(* IEC 61131-3 sources: daoli-st-library/DL_Process (part 63) *)

(* ---- FB_DL_ChamberSeasoningTrack.st ---- *)
(*==============================================================================
 * 组件名称 (Component)  : FB_DL_ChamberSeasoningTrack
 * 所属子库 (Sublibrary) : DL_Process
 * 当前版本 (Version)    : 1.0.0
 * 组件分类 (Category)   : 功能块（FUNCTION_BLOCK）· 腔体 seasoning 台账与放行判定
 * 兼容性   (Platform)   : CODESYS 3.5 / TwinCAT 3 / 汇川 InoProShop / Schneider Machine Expert
 *                         仅依赖 Standard.library（R_TRIG / LEN / LEFT / ABS / MIN / MAX / LIMIT），零厂商方言
 * 接口依赖 (Depends)    : E_DL_Ne107Status —— 唯一属主为 DL_Device 子库的契约件
 *                         I_DL_DeviceHealth（R13 泳道 A1）。本文件只引用成员，不重定义枚举体。
 * 功能描述 (Function)   : seasoning（腔体调机）片数 + 膜厚台账 + 放行判定。每片完成后累计
 *                         片数、累计工艺时长、膜厚均值与趋势；**双判据**（片数达标 **且** 时长
 *                         达标）才放行；连续越窗自动降级 eNotReady；配方名只作标签与校验键。
 * 边界     (Boundary)   : ① **不做配方存储** —— sRecipeName 只作为标签与校验键传入，配方本体
 *                         归 FB_DL_RecipeManager；② **不做膜厚测量** —— 膜厚与均匀性由量测机台
 *                         引脚注入；③ 不做 SPC 判异（只做越窗计数与连续计数）；④ 不做 MES 上报。
 * 分层声明 (Layer)      : 工艺层（DL_Process）。零全局变量表引用、零外部变量声明、零物理 IO。
 * 段序     (Segments)   : 段1 实例无条件刷新 → 段2 复位通道（CASE 前，R39）→ 段3 配方标签闸门
 *                         （R37 显式截断）与参数钳位 → 段4 单片完成受理（R24/R25/R44）→
 *                         段5 状态机 → 段6 码位单一优先级链 → 段7 出口钳位与保持重写。
 * 枚举映射表 (R31)      : eIdle(0)→标签 0｜eTracking(10)→标签 10｜eQualified(20)→标签 20｜
 *                         eNotReady(30)→标签 30｜eFault(99)→标签 99。每个成员有且仅有一个
 *                         显式标签，ELSE 只接脏值（02FB）。
 * 单拍标志清单 (R25)    : bWaferDone —— 预清零点：段1 每拍被实例输出覆盖；置位点：段1
 *                         `_bWaferReq := _fbTrigWafer.Q AND (NOT _bWaferConsumed)`；自清点：
 *                         段4 消费时置 `_bWaferConsumed := TRUE`，bWaferDone 回 FALSE 即解除。
 *                         bReset —— 预清零点：段1 覆盖 _bResetEdge；置位点：段1 实例调用；
 *                         自清点：紧随实例调用的 _bResetEdge 赋值行。
 * 保持位清单 (R27)      : bRelease 逐拍由 _bReleaseLatched 重写；eQualify 逐拍由 _eState 映射；
 *                         nCount / nNgCount / tAccum / fThickAvg / fThickSlope 逐拍由内部
 *                         台账量重写并夹域。复位沿清台账并递增轮次号。
 * 定时器清单 (R40)      : 无 TON/TOF 实例。工艺时长由引脚 tProcessTime 累加（台账语义），
 *                         不存在跨段恒真的定时输入；片数与时长的「达标」判据均为纯比较式。
 * 三元一致表 (R35)      : 片数目标守卫 1~10000 / 封顶 10000 / 判据 `>=`｜
 *                         连续越窗阈守卫 1~10 / 封顶 10 / 判据 `>=`｜
 *                         膜厚容差守卫 0.5~50 % / 封顶 50 / 判据 `>`（越窗）。
 * 镜像量清单 (R38)      : sRecipeName 的长度经 LEN 一次锁存为 _nNameLen，截断判定与登记
 *                         全部读该锁存量，绝不二次取长度；fThickness 与 fUniformity 在段4
 *                         单次锁存后参与全部判据。
 * 开源溯源 (Origin)     : 原创实现（参考 SEMI/半导体厂务公开的 seasoning 台账惯例，以及
 *                         ISA-88 公开的批次/相语义，T2-8 只借「批次台账 + 放行」的组织形态；
 *                         配方名仅作标签、台账只做累计与双判据）。ISA-88 为公开标准条款，
 *                         不声称「符合 ISA-88」；实现、码位、引脚契约 100% 本库独立设计，
 *                         clean-room 编写，未复制任何源码行。许可证说明：无代码借鉴对象，
 *                         本文件为本库原创，随本库许可证发布。
 * 验收向量 (Acceptance) :
 *   V1 25 片、每片 24 min、膜厚 100 ± 2 nm（目标 100、容差 5 %）→ tAccum = 10 h、
 *      eQualified、bRelease = TRUE。
 *   V2（双判据）25 片但每片 10 min（总 4.17 h < 10 h）→ 16#0005_01CD、仍 eTracking、
 *      bRelease = FALSE。
 *   V3（V-A 缺失键）sRecipeName = '' → 16#0005_02F9 锁存、bRelease 强制 FALSE
 *      （安全侧：台账不可信不得放行）。
 *   V4（V-B 串上限，R37）sRecipeName 传 40 字符（超 STRING(32)）→ 入口判 LEN 后置
 *      16#0005_01CE，按截断后的名字登记台账，**不得**依赖赋值隐式截断后静默使用。
 *   V5（V-D 复位首拍）bReset 后 nCount = 0、tAccum = T#0S、nRoundId + 1、bRelease = FALSE；
 *      **不得**保留上一轮 fThickSlope 的首片基准（R41：恢复不重头）。
 * 偏离留档 (Deviation)  :
 *   ① sRecipeName 引脚类型由 STRING(32) 提升为 STRING(80)：若按 STRING(32) 声明，超长截断
 *      会发生在**调用方赋值**那一行，本件永远看不到长度越限，01CE 成为死码 —— 这正是 R37
 *      要消灭的「静默截断」。提升到 STRING(80) 后由本件判 LEN、显式置码、按截断名登记，
 *      登记缓冲仍为 STRING(32)（_sRecipeTag），行为与规格 V4 一致。
 *   ② 工艺时长用 tProcessTime 累加而非墙钟：一台上位机可能同时跟踪多条腔体，墙钟会把
 *      「等待/待机」算进 seasoning 时长；引脚注入的工艺耗时才是台账口径。
 *   ③ 越窗判据取「膜厚相对偏差 > fThickTol 或 均匀性 > fUnifLimit」的**并集**：均匀性越限
 *      同样是「膜质未稳」的证据，只盯膜厚会漏掉「厚度对但均匀性崩」的片子。
 *   ④ 量测值非有限/越域并入 16#0005_02FA：规格故障表只给三个码，量测值不可信属于
 *      「台账数据源坏了」，与计数溢出同属「台账不可继续累加」的语义，故共用该码；
 *      不发生任何累加（本片不入账），也不会放行。
 * 修订历史 (Revision)   :
 *   2026-11-15  v1.0.0  首版入库（Round 13 · 泳道 C · DL_Process 第 25 件）
 *============================================================================*)

(*-----------------------------------------------------------------------------
 * 枚举: E_DL_SeasonState（归属 FB_DL_ChamberSeasoningTrack，同文件发布）
 *----------------------------------------------------------------------------*)
TYPE E_DL_SeasonState :
(
    eIdle      := 0,    // 空闲：未使能或参数未就绪 / Idle, disabled or parameters not ready
    eTracking  := 10,   // 台账中：逐片累计，双判据未齐 / Tracking, accumulating wafers
    eQualified := 20,   // 已放行：片数与时长双达标 / Qualified, both criteria met
    eNotReady  := 30,   // 不具备放行条件：连续越窗降级 / Not ready, consecutive out-of-window wafers
    eFault     := 99    // 故障：配方键缺失或计数溢出 / Fault, missing recipe key or counter overflow
) UINT;
END_TYPE

FUNCTION_BLOCK FB_DL_ChamberSeasoningTrack
VAR_INPUT
    bEnable       : BOOL;                   // 使能（Enable），FALSE = 冻结台账与放行；复位通道不受其屏蔽 / Enable, FALSE freezes the ledger
    bReset        : BOOL;                   // 复位（Reset），上升沿清台账并重开新一轮 / Rising edge clears the ledger and opens a new round
    bWaferDone    : BOOL;                   // 单片完成（One-shot wafer done），上升沿受理（R24）/ One-shot wafer done, rising edge only
    fThickness    : REAL;                   // 本片膜厚（Wafer thickness）[nm]，域 0~10000 / Wafer thickness [nm], 0 to 10000
    fUniformity   : REAL;                   // 本片均匀性（Uniformity）[%]，域 0~100 / Uniformity [%], 0 to 100
    sRecipeName   : STRING(80);             // 配方名标签（Recipe tag），域非空，超 32 字符显式截断并置码（偏离留档①）/ Recipe tag, truncated explicitly
    fThickTarget  : REAL;                   // 膜厚目标（Thickness target）[nm]，域 >0 / Thickness target [nm], must be positive
    fThickTol     : REAL := 5.0;            // 膜厚相对容差（Thickness tolerance）[%]，域 0.5~50，默认 5.0 / Thickness tolerance [%]
    fUnifLimit    : REAL := 3.0;            // 均匀性上限（Uniformity limit）[%]，域 0.1~20，默认 3.0 / Uniformity limit [%]
    nCountTarget  : INT := 25;              // 片数目标（Wafer count target）[片]，域 1~10000，默认 25 / Wafer count target [pcs]
    tTimeTarget   : TIME := T#10H;          // 工艺时长目标（Process time target），域 1 min~1000 h，默认 10 h / Process time target
    nConsecNgLimit : INT := 2;              // 连续越窗降级阈值（Consecutive out-of-window limit）[片]，域 1~10，默认 2 / Consecutive limit [pcs]
    tProcessTime  : TIME;                   // 本片工艺耗时（Process time of this wafer），由上层引脚注入 / Process time injected by the caller
END_VAR

VAR_OUTPUT
    nCount        : INT;                    // 已 seasoning 片数（Seasoned wafer count）[片]，逐拍重写 / Seasoned wafer count [pcs]
    nNgCount      : INT;                    // 越窗片数（Out-of-window wafer count）[片]，逐拍重写 / Out-of-window wafer count [pcs]
    tAccum        : TIME;                   // 累计工艺时长（Accumulated process time），逐拍重写 / Accumulated process time
    fThickAvg     : REAL;                   // 膜厚均值（Mean thickness）[nm]，逐拍重写 / Mean thickness [nm]
    fThickSlope   : REAL;                   // 膜厚趋势（Thickness trend）[nm/片]，首末差除以片数差 / Thickness trend [nm/pc]
    bRelease      : BOOL;                   // 放行（Release），保持语义（R27）/ Release, held
    eQualify      : E_DL_SeasonState;       // 判定状态（Qualification state），逐拍重写 / Qualification state
    nRoundId      : UINT;                   // 本轮编号（Round id），复位递增，供 MES 对齐 / Round id, incremented on reset
    eHealth       : E_DL_Ne107Status;       // 健康态（NE107 health），引用属主 A1 的枚举 / NE107 health, owned by A1
    uDiagCode     : UDINT;                  // 诊断码（Diagnostic code），本拍单一优先级链输出 / Diagnostic code, single priority chain
    uErrorId      : UDINT;                  // 故障码（Error code），仅故障级码，0 = 无故障 / Fault-level code, 0 = no fault
    bError        : BOOL;                   // 故障标志（Error），仅故障级码置位 / TRUE only for fault-level codes
END_VAR

VAR
    _eState       : E_DL_SeasonState := E_DL_SeasonState.eIdle;    // 内部状态（Internal state）/ Internal state value
    _bWaferReq    : BOOL;                   // 单片完成单拍请求（Wafer done request）/ Wafer done one-shot request
    _bWaferConsumed : BOOL;                 // 单片完成已消费（Wafer consumed flag）/ Wafer consumed flag
    _bResetEdge   : BOOL;                   // 复位沿单拍标志（Reset one-shot flag）/ Reset one-shot flag
    _uFaultCode   : UDINT;                  // 本拍故障级码（Fault-level code this scan）/ Fault-level code of this scan
    _uFaultLatched : UDINT;                 // 故障码锁存（Latched fault code），仅复位清除 / Latched fault code, reset only
    _uInfoCode    : UDINT;                  // 本拍信息级码（Info-level code this scan）/ Info-level code of this scan
    _bFaultCond   : BOOL;                   // 故障条件（Fault condition）/ Fault condition flag
    _sRecipeTag   : STRING(32);             // 台账登记的配方标签（Registered recipe tag），截断后 32 字符 / Recipe tag after truncation
    _nNameLen     : INT;                    // 配方名长度（Recipe name length）[字符]，一次锁存（R38）/ Recipe name length, latched once
    _bTruncFlag   : BOOL;                   // 截断发生标志（Truncation flag），R37 显式置位 / Truncation flag, set explicitly (R37)
    _bKeyOk       : BOOL;                   // 配方键与目标合法（Key and target valid）/ Key and target valid
    _fThickSnap   : REAL;                   // 膜厚快照（Thickness snapshot）[nm]，单次锁存 / Thickness snapshot [nm]
    _fUnifSnap    : REAL;                   // 均匀性快照（Uniformity snapshot）[%]，单次锁存 / Uniformity snapshot [%]
    _fTolEff      : REAL;                   // 生效膜厚容差（Effective thickness tolerance）[%] / Effective thickness tolerance [%]
    _fUnifLimEff  : REAL;                   // 生效均匀性上限（Effective uniformity limit）[%] / Effective uniformity limit [%]
    _nCountTgtEff : INT;                    // 生效片数目标（Effective count target）[片] / Effective count target [pcs]
    _nConsecEff   : INT;                    // 生效连续越窗阈（Effective consecutive limit）[片] / Effective consecutive limit [pcs]
    _tTimeTgtEff  : TIME;                   // 生效时长目标（Effective time target）/ Effective time target
    _nCountInt    : INT;                    // 内部片数台账（Internal wafer count）[片] / Internal wafer count [pcs]
    _nNgInt       : INT;                    // 内部越窗片数（Internal out-of-window count）[片] / Internal out-of-window count [pcs]
    _nConsecNg    : INT;                    // 当前连续越窗片数（Current consecutive out-of-window count）[片] / Current consecutive count [pcs]
    _tAccumInt    : TIME;                   // 内部累计时长（Internal accumulated time）/ Internal accumulated time
    _fThickSum    : REAL;                   // 膜厚累加（Thickness sum）[nm] / Thickness sum [nm]
    _fThickFirst  : REAL;                   // 首片膜厚（First wafer thickness）[nm]，趋势基准 / First wafer thickness [nm]
    _fThickLast   : REAL;                   // 末片膜厚（Last wafer thickness）[nm] / Last wafer thickness [nm]
    _bFirstSet    : BOOL;                   // 首片基准已装（First sample recorded）/ First sample recorded flag
    _fDevPct      : REAL;                   // 膜厚相对偏差（Relative thickness deviation）[%] / Relative thickness deviation [%]
    _bOutWin      : BOOL;                   // 本片越窗（Out of window this wafer）/ Out of window this wafer
    _bReleaseLatched : BOOL;                // 放行锁存（Release latch），复位清除 / Release latch, reset only
    _nRoundIdInt  : UINT;                   // 内部轮次号（Internal round id），复位递增 / Internal round id, incremented on reset
    _bCountOk     : BOOL;                   // 片数达标（Count criterion met）/ Count criterion met
    _bTimeOk      : BOOL;                   // 时长达标（Time criterion met）/ Time criterion met
    _fbTrigWafer  : R_TRIG;                 // 单片完成上升沿（Wafer done rising edge）/ Wafer done rising edge
    _fbTrigReset  : R_TRIG;                 // 复位上升沿（Reset rising edge）/ Reset rising edge
END_VAR

VAR CONSTANT
    DL_SEA_NAME_MAX   : INT  := 32;          // 配方标签登记宽度（Registered tag width）[字符]，与 STRING(32) 一致 / Registered tag width
    DL_SEA_REAL_MAX   : REAL := 3.4E38;      // 单精度有限值判据幅值（Finite magnitude bound）/ Finite bound for REAL inputs
    DL_SEA_EPS        : REAL := 1.0E-6;      // 浮点防零容差（Divide-guard epsilon）/ Float divide-guard epsilon
    DL_SEA_THICK_MAX  : REAL := 10000.0;     // 膜厚输入域上限（Thickness input bound）[nm] / Thickness input bound [nm]
    DL_SEA_UNIF_MAX   : REAL := 100.0;       // 均匀性输入域上限（Uniformity input bound）[%] / Uniformity input bound [%]
    DL_SEA_TOL_LO     : REAL := 0.5;         // 膜厚容差下限（Tolerance lower clamp）[%] / Tolerance lower clamp [%]
    DL_SEA_TOL_HI     : REAL := 50.0;        // 膜厚容差上限（Tolerance upper clamp）[%] / Tolerance upper clamp [%]
    DL_SEA_UNIFL_LO   : REAL := 0.1;         // 均匀性上限下限（Uniformity limit lower clamp）[%] / Uniformity lower clamp [%]
    DL_SEA_UNIFL_HI   : REAL := 20.0;        // 均匀性上限上限（Uniformity limit upper clamp）[%] / Uniformity upper clamp [%]
    DL_SEA_CNT_LO     : INT  := 1;           // 片数目标下限（Count target lower clamp）[片] / Count target lower clamp [pcs]
    DL_SEA_CNT_HI     : INT  := 10000;       // 片数目标上限（Count target upper clamp）[片] / Count target upper clamp [pcs]
    DL_SEA_CONS_LO    : INT  := 1;           // 连续阈下限（Consecutive limit lower clamp）[片] / Consecutive limit lower clamp [pcs]
    DL_SEA_CONS_HI    : INT  := 10;                 // 连续阈上限（Consecutive limit upper clamp）[片] / Consecutive limit upper clamp [pcs]
    DL_SEA_CNT_OVF    : INT  := 30000;       // 片数台账溢出阈（Count overflow threshold）[片] / Count overflow threshold [pcs]
    DL_SEA_TIME_OVF   : TIME := T#40D;       // 时长台账溢出阈（Time overflow threshold）[ms] / Time overflow threshold
    DL_SEA_TIME_MIN   : TIME := T#1M;        // 时长目标下限（Time target lower clamp）/ Time target lower clamp
    DL_SEA_TIME_MAX   : TIME := T#1000H;     // 时长目标上限（Time target upper clamp）/ Time target upper clamp
    DL_SEA_PCT        : REAL := 100.0;       // 百分比换算（Percent scale）[-] / Percent scale
    DL_SEA_ERR_KEY    : UDINT := 16#0005_02F9; // 0005_02F9 配方名为空或膜厚目标非正【故障级】/ Missing recipe or target, fault level
    DL_SEA_ERR_OVF    : UDINT := 16#0005_02FA; // 0005_02FA 片数或时长台账溢出【故障级】/ Counter overflow, fault level
    DL_SEA_ERR_STATE  : UDINT := 16#0005_02FB; // 0005_02FB 非法状态兜底【故障级】/ Illegal state fallback, fault level
    DL_SEA_INFO_SINGLE : UDINT := 16#0005_01CB; // 0005_01CB 单片越窗但未连续【信息级】/ Single out-of-window wafer, info level
    DL_SEA_INFO_CONS  : UDINT := 16#0005_01CC; // 0005_01CC 连续越窗达阈值降级【信息级】/ Consecutive limit reached, info level
    DL_SEA_INFO_TIME  : UDINT := 16#0005_01CD; // 0005_01CD 片数达标但时长未达标【信息级】/ Count reached, time pending, info level
    DL_SEA_INFO_TRUNC : UDINT := 16#0005_01CE; // 0005_01CE 配方名超 32 字符已显式截断【信息级】/ Recipe tag truncated explicitly, info level
END_VAR

// ============================================================================
// 段 1｜实例无条件周期刷新（R7/0.5：严禁置于 IF / CASE 分支内）
//      Unconditional per-cycle refresh of every instance (R7/0.5)
// ============================================================================
_fbTrigWafer(CLK := bWaferDone);                // 单片完成上升沿（Wafer done rising edge）
_bWaferReq := _fbTrigWafer.Q AND (NOT _bWaferConsumed);    // 单拍请求（R25 置位点）
_fbTrigReset(CLK := bReset);                    // 复位上升沿（Reset rising edge）
_bResetEdge := _fbTrigReset.Q;                  // 复位单拍标志紧随实例赋值（R25 自清点）

// 本拍码与条件预置（每拍重算；故障码以上拍锁存续用）
// Per-scan preset of codes and conditions, the fault code is carried from the latch
_uFaultCode := _uFaultLatched;                  // 故障码续用（Carry the latched fault code）
_uInfoCode  := 16#0000_0000;                    // 信息级码预清零（Info code preset to zero）
_bFaultCond := FALSE;                           // 故障条件预清零（Fault condition preset FALSE）
_bKeyOk     := FALSE;                           // 配方键闸门预置未通过（Key gate preset closed）
_bOutWin    := FALSE;                           // 越窗标志预置假（Out-of-window preset FALSE）

// 单片完成消费标志解除：输入回落即允许下一片（R25 生命周期闭环）
// Release the wafer consumption flag once the input falls
IF NOT bWaferDone THEN
    _bWaferConsumed := FALSE;                   // 允许下一次上升沿（Next rising edge accepted）
END_IF

// ============================================================================
// 段 2｜复位通道（R39：置于 CASE 之前，且不被掉使能分支屏蔽）
//      Reset path, before CASE and never masked by the disable branch
// ============================================================================
IF _bResetEdge THEN
    _nCountInt    := 0;                         // 片数台账清零（Wafer count cleared）
    _nNgInt       := 0;                         // 越窗片数清零（Out-of-window count cleared）
    _nConsecNg    := 0;                         // 连续越窗计数清零（Consecutive count cleared）
    _tAccumInt    := T#0S;                      // 累计时长清零（Accumulated time cleared）
    _fThickSum    := 0.0;                       // 膜厚累加清零（Thickness sum cleared）
    _fThickFirst  := 0.0;                       // 首片基准清除（First-sample basis cleared）
    _fThickLast   := 0.0;                       // 末片值清除（Last-sample value cleared）
    _bFirstSet    := FALSE;                     // 首片基准标志清除（First-sample flag cleared，R41）
    _bReleaseLatched := FALSE;                  // 放行锁存清除（Release latch cleared）
    _bTruncFlag   := FALSE;                     // 截断标志清除（Truncation flag cleared）
    _nRoundIdInt  := _nRoundIdInt + UINT#1;     // 轮次递增进位（Round id incremented）
    _uFaultLatched := 16#0000_0000;             // 故障码锁存清除（Latched fault code cleared）
    _uFaultCode   := 16#0000_0000;              // 本拍故障码清空，防止段6 重新锁存旧码（Clear this scan code）
    IF _eState = E_DL_SeasonState.eFault THEN
        _eState := E_DL_SeasonState.eIdle;      // 故障态回空闲（Fault state back to idle）
        _bFaultCond := FALSE;                   // 故障条件清除（Fault condition cleared）
    ELSIF _eState = E_DL_SeasonState.eQualified THEN
        _eState := E_DL_SeasonState.eTracking;  // 已放行轮次复位后重开台账（New round after a qualified round）
    ELSIF _eState = E_DL_SeasonState.eNotReady THEN
        _eState := E_DL_SeasonState.eTracking;  // 降级轮次复位后重开台账（New round after a degraded round）
    END_IF
END_IF

// ============================================================================
// 段 3｜配方标签闸门（R37：先判长度、显式置码、按截断名登记）与参数钳位
//      Recipe tag gate: length first, explicit code, then register the truncated tag
// ============================================================================
_nNameLen := LEN(sRecipeName);                  // 长度一次锁存（R38：此后全部判据读该值）
IF _nNameLen > DL_SEA_NAME_MAX THEN
    _sRecipeTag := LEFT(sRecipeName, DL_SEA_NAME_MAX);   // 按宽度取前缀后写回登记缓冲（预判后写，非回夹）
    _bTruncFlag := TRUE;                        // 截断标志显式置位（R37 核心：不静默）
    _uInfoCode  := DL_SEA_INFO_TRUNC;           // 0005_01CE 配方名超长已截断【信息级】/ Recipe tag truncated
ELSE
    _sRecipeTag := sRecipeName;                 // 未超长按原名登记（Register the tag as-is）
END_IF

IF _nNameLen = 0 THEN
    _bFaultCond := TRUE;                        // 配方键缺失（Missing recipe key）
    _uFaultCode := DL_SEA_ERR_KEY;              // 0005_02F9 配方名为空【故障级】/ Missing recipe, fault level
ELSIF (NOT (fThickTarget >= DL_SEA_EPS)) OR (fThickTarget > DL_SEA_THICK_MAX) THEN
    _bFaultCond := TRUE;                        // 膜厚目标非正或越域（Target not positive or out of domain）
    _uFaultCode := DL_SEA_ERR_KEY;              // 0005_02F9 膜厚目标非法【故障级】/ Illegal target, fault level
ELSE
    _bKeyOk := TRUE;                            // 键与目标合法（Key and target valid）
END_IF

// 参数域钳位（R35：守卫、封顶与判据同向）
// Parameter clamping so that guard, ceiling and comparison stay in step (R35)
_fTolEff      := LIMIT(DL_SEA_TOL_LO, fThickTol, DL_SEA_TOL_HI);            // 膜厚容差 0.5~50 %（Tolerance clamped）
_fUnifLimEff  := LIMIT(DL_SEA_UNIFL_LO, fUnifLimit, DL_SEA_UNIFL_HI);       // 均匀性上限 0.1~20 %（Uniformity limit clamped）
_nCountTgtEff := LIMIT(DL_SEA_CNT_LO, nCountTarget, DL_SEA_CNT_HI);         // 片数目标 1~10000（Count target clamped）
_nConsecEff   := LIMIT(DL_SEA_CONS_LO, nConsecNgLimit, DL_SEA_CONS_HI);     // 连续阈 1~10（Consecutive limit clamped）
_tTimeTgtEff := tTimeTarget;                    // 时长目标取引脚值（Time target taken from the pin）
IF _tTimeTgtEff < DL_SEA_TIME_MIN THEN
    _tTimeTgtEff := DL_SEA_TIME_MIN;            // 时长目标下限钳位（Time target lower clamp）
ELSIF _tTimeTgtEff > DL_SEA_TIME_MAX THEN
    _tTimeTgtEff := DL_SEA_TIME_MAX;            // 时长目标上限钳位（Time target upper clamp）
END_IF

// ============================================================================
// 段 4｜单片完成受理（R24/R25；R44 清码点绑定新片起点）
//      Wafer completion acceptance, info codes cleared at each wafer start (R44)
// ============================================================================
IF _bWaferReq AND (NOT _bWaferConsumed) AND (_eState = E_DL_SeasonState.eTracking) AND _bKeyOk THEN
    _bWaferConsumed := TRUE;                    // 消费单片沿（Wafer edge consumed）
    _uInfoCode      := 16#0000_0000;            // 新片起点清信息码（R44：清码点绑定新片起点）
    _fThickSnap     := fThickness;              // 膜厚快照（Thickness snapshot）
    _fUnifSnap      := fUniformity;             // 均匀性快照（Uniformity snapshot）

    IF (NOT (_fThickSnap >= 0.0 AND _fThickSnap <= DL_SEA_THICK_MAX))
    OR (NOT (_fUnifSnap >= 0.0 AND _fUnifSnap <= DL_SEA_UNIF_MAX)) THEN
        _bFaultCond := TRUE;                    // 量测值非有限或越域（Non-finite or out-of-domain measurement）
        _uFaultCode := DL_SEA_ERR_OVF;          // 0005_02FA 量测值非法并入溢出码【故障级】/ Illegal measurement folded in
    ELSE
        _nCountInt := _nCountInt + 1;           // 片数 +1（Wafer counted）
        _fThickSum := _fThickSum + _fThickSnap; // 膜厚累加（Thickness accumulated）
        _fThickLast := _fThickSnap;             // 末片膜厚（Last wafer thickness）
        IF NOT _bFirstSet THEN
            _fThickFirst := _fThickSnap;        // 首片基准只在首片装一次（First-sample basis once）
            _bFirstSet   := TRUE;               // 基准已装（Basis recorded）
        END_IF
        _tAccumInt := _tAccumInt + tProcessTime;    // 累计工艺时长（Process time accumulated）

        // 越窗判据：膜厚相对偏差 或 均匀性越限（偏离留档③）
        //     Out-of-window when the thickness deviation or the uniformity exceeds its limit
        _fDevPct := ABS(_fThickSnap - fThickTarget) / fThickTarget * DL_SEA_PCT;    // 相对偏差（Relative deviation）
        IF (_fDevPct > _fTolEff) OR (_fUnifSnap > _fUnifLimEff) THEN
            _bOutWin := TRUE;                   // 本片越窗（Out of window）
        END_IF

        IF _bOutWin THEN
            _nNgInt    := _nNgInt + 1;          // 越窗片数 +1（Out-of-window counted）
            _nConsecNg := _nConsecNg + 1;       // 连续越窗 +1（Consecutive count increments）
            IF _nConsecNg >= _nConsecEff THEN
                _uInfoCode := DL_SEA_INFO_CONS; // 0005_01CC 连续越窗达阈值降级【信息级】/ Consecutive limit reached
            ELSE
                _uInfoCode := DL_SEA_INFO_SINGLE;   // 0005_01CB 单片越窗但未连续【信息级】/ Single out-of-window wafer
            END_IF
        ELSE
            _nConsecNg := 0;                    // 未越窗则连续计数清零（Consecutive count resets）
        END_IF

        // 台账溢出守卫（R35：守卫 30000 片 / 40 天，判据 >=）
        //     Ledger overflow guard
        IF (_nCountInt >= DL_SEA_CNT_OVF) OR (_tAccumInt >= DL_SEA_TIME_OVF) THEN
            _bFaultCond := TRUE;                // 台账溢出（Ledger overflow）
            _uFaultCode := DL_SEA_ERR_OVF;      // 0005_02FA 台账溢出【故障级】/ Ledger overflow, fault level
        END_IF
    END_IF
END_IF

// 双判据（片数达标 且 时长达标）：片数达标而时长未达标时只给信息码，不放行
// Dual criteria: the count alone never releases the chamber
_bCountOk := _nCountInt >= _nCountTgtEff;       // 片数判据（Count criterion）
_bTimeOk  := _tAccumInt >= _tTimeTgtEff;        // 时长判据（Time criterion）
IF _bCountOk AND (NOT _bTimeOk) THEN
    _uInfoCode := DL_SEA_INFO_TIME;             // 0005_01CD 片数达标但时长未达标【信息级】/ Count reached, time pending
END_IF

// ============================================================================
// 段 5｜状态机（ENUM + CASE，含 ELSE 非法状态兜底）
//      State machine with an explicit ELSE fallback
// ============================================================================
IF _bFaultCond THEN
    _bReleaseLatched := FALSE;                  // 安全侧：台账不可信时强制撤销放行（Safety: release revoked on any fault）
    _eState := E_DL_SeasonState.eFault;         // 故障条件优先于状态机（Fault outranks the machine）
END_IF

// 掉使能冻结分支：显式排除故障态（R39 合法写法①），复位通道仍可从故障态退出
// Disable branch explicitly excludes the fault state so the reset path still works
IF (NOT bEnable) AND (_eState <> E_DL_SeasonState.eFault) THEN
    _eState := E_DL_SeasonState.eIdle;          // 冻结回空闲（Freeze back to idle）
END_IF

CASE _eState OF

    E_DL_SeasonState.eIdle: // 空闲：等键与目标就绪
        IF bEnable AND _bKeyOk AND (NOT _bFaultCond) THEN
            _eState := E_DL_SeasonState.eTracking;  // 门票就绪进台账（Enter tracking）
        END_IF

    E_DL_SeasonState.eTracking: // 台账中：双判据 / 连续越窗降级
        IF _bCountOk AND _bTimeOk THEN
            _bReleaseLatched := TRUE;           // 双判据齐：放行（Releases the chamber）
            _eState := E_DL_SeasonState.eQualified; // 进已放行（Enter qualified）
        ELSIF _nConsecNg >= _nConsecEff THEN
            _bReleaseLatched := FALSE;          // 降级：撤销放行（Degraded, release revoked）
            _eState := E_DL_SeasonState.eNotReady;  // 进不具备放行条件（Enter not ready）
        END_IF

    E_DL_SeasonState.eQualified: // 已放行：结论逐拍在段7 重写（R27），本分支只保留标签
        // 结论保持由段7 逐拍重写承担，此处保留空标签与原因注释（R31）
        // The held verdict is rewritten in segment 7, so this label stays empty (R31)

    E_DL_SeasonState.eNotReady: // 不具备放行条件：等复位重开一轮
        // 复位通道位于 CASE 之前（段2），此处保留空标签与原因注释（R31/R41）
        // Reset happens in segment 2, so this label stays empty (R31/R41)

    E_DL_SeasonState.eFault: // 故障：等复位沿（段2）
        // 复位通道位于 CASE 之前，此分支无需动作（R39）
        // The reset path sits before CASE, so no action is needed here (R39)

    ELSE // 兜底：非法状态
        _uFaultCode := DL_SEA_ERR_STATE;        // 0005_02FB 非法状态兜底【故障级】/ Illegal state fallback
        _bFaultCond := TRUE;                    // 置故障条件（Raise the fault condition）
        _eState     := E_DL_SeasonState.eFault; // 强制回故障态（Force the fault state）
END_CASE

// ============================================================================
// 段 6｜码位单一优先级链（全拍只写一次，信息级不置 bError）
//      Single priority chain for the codes, written once per scan
// ============================================================================
IF _uFaultCode <> 16#0000_0000 THEN
    _uFaultLatched := _uFaultCode;              // 故障码锁存（Latched until reset）
    uErrorId  := _uFaultCode;                   // 故障级码优先（Fault-level code wins）
    uDiagCode := _uFaultCode;                   // 诊断码同源（Diagnostic code mirrors the fault）
    bError    := TRUE;                          // 故障标志置位（Error flag raised）
ELSIF _uInfoCode <> 16#0000_0000 THEN
    uErrorId  := 16#0000_0000;                  // 信息级不占故障码（Info level leaves the fault code empty）
    uDiagCode := _uInfoCode;                    // 诊断码取信息级码（Diagnostic code takes the info code）
    bError    := FALSE;                         // 信息级不置故障位（Info level never raises the error flag）
ELSE
    uErrorId  := 16#0000_0000;                  // 无码（No code）
    uDiagCode := 16#0000_0000;                  // 无码（No code）
    bError    := FALSE;                         // 无故障（No error）
END_IF

// ============================================================================
// 段 7｜出口钳位与保持语义重写（R27/R43；台账量逐拍重写，绝不靠进入那一拍）
//      Output clamping and held-semantics rewrite (R27/R43)
// ============================================================================
nCount    := LIMIT(0, _nCountInt, DL_SEA_CNT_OVF);      // 片数夹进 0~30000（Count clamped）
nNgCount  := LIMIT(0, _nNgInt, DL_SEA_CNT_OVF);         // 越窗片数夹进 0~30000（Out-of-window clamped）
tAccum    := _tAccumInt;                                // 累计时长逐拍重写（Accumulated time rewritten）
IF _nCountInt > 0 THEN
    fThickAvg := _fThickSum / INT_TO_REAL(_nCountInt);  // 膜厚均值（Mean thickness），除零已由计数守卫
ELSE
    fThickAvg := 0.0;                                   // 无片时均值 0（Zero mean without wafers）
END_IF
IF (_nCountInt >= 2) AND _bFirstSet THEN
    fThickSlope := (_fThickLast - _fThickFirst) / INT_TO_REAL(_nCountInt - 1);  // 首末差/片数差（Trend per wafer）
ELSE
    fThickSlope := 0.0;                                 // 单片或未装基准时趋势 0（Zero trend before a basis exists）
END_IF
bRelease  := _bReleaseLatched;                          // 放行逐拍重写（Release rewritten every scan）
eQualify  := _eState;                                   // 判定状态逐拍重写（Qualification state rewritten）
nRoundId  := _nRoundIdInt;                              // 轮次号逐拍重写（Round id rewritten every scan）

// 健康态仲裁（引用属主 A1 的四态语言）
// Health arbitration mapped onto the A1 health language
IF _eState = E_DL_SeasonState.eFault THEN
    eHealth := E_DL_Ne107Status.eFailure;       // 故障：台账不可信（Failure）
ELSIF NOT bEnable THEN
    eHealth := E_DL_Ne107Status.eUnknown;       // 未知：未使能（Unknown）
ELSIF _eState = E_DL_SeasonState.eNotReady THEN
    eHealth := E_DL_Ne107Status.eMaintenanceReq;    // 需维护：连续越窗，需重新调机（Maintenance required）
ELSIF _bTruncFlag THEN
    eHealth := E_DL_Ne107Status.eOutOfSpec;     // 越规：配方键被截断，台账对齐风险（Out of spec）
ELSIF _eState = E_DL_SeasonState.eQualified THEN
    eHealth := E_DL_Ne107Status.eOk;            // 正常：已放行（OK, released）
ELSE
    eHealth := E_DL_Ne107Status.eOk;            // 正常：台账进行中（OK, tracking）
END_IF

END_FUNCTION_BLOCK

(* ---- FB_DL_CipCleaningSeq.st ---- *)
(*==============================================================================
 * 组件名称 (Component)  : FB_DL_CipCleaningSeq
 * 所属子库 (Sublibrary) : DL_Process
 * 当前版本 (Version)    : 1.0.1
 * 兼容性 (Platform)   : CODESYS 3.5 / TwinCAT 3 / 汇川 InoProShop / Machine Expert
 *                         仅依赖 Standard.library（TON / R_TRIG），零厂商方言
 * 分类     (Category)   : 工艺段功能块（Function Block · CIP 原位清洗六相顺控）
 * 功能简述 (Function)   : CIP 原位清洗六相顺控：预冲洗 → 碱洗 → 中间冲洗 →
 *                         酸洗 → 终冲洗 → 消毒。核心纪律：相位计时受 TACT 联
 *                         锁暂停（温度/电导率/流量不达标不计时）；终冲洗以回
 *                         液电导率判终点（最长延时兜底）；回路就绪门控；换相
 *                         停泵间隔防混液；中止即排空隔离并失去清洁许可；偏差
 *                         计数供审计。本块不实现阀门矩阵/混流防护的物理设计
 *                         （属机械与管路设计），仅做就绪门控与指令编排。
 * 首扫说明 (Init note)  : 顺序型组件但全部状态由指令沿/电平驱动，免首扫
 *                         （R23/公约 0.1），无 bInit。
 * 公约遵循 (Convention) : 0.2/R21 bError 仅故障级码置位；0.4 双语同行注释；
 *                         0.5/R7 八实例（R_TRIG×2/TON×6）主体最前部无条件刷
 *                         新；0.7/R15 故障锁存仅复位路径清码；0.10 定时基准
 *                         由引脚给（tCycle 增补引脚，泳道 A 同款公共约定）；
 *                         0.14 数组存取先判域（所有相位索引先判 < 上限）、
 *                         FOR 有界（无 WHILE）、非有限值防御；0.15 温度 ℃、
 *                         电导率 mS/cm、流量 m³/h，同块不混用；0.16 无魔法
 *                         数；0.17 终结符成对 ✓；0.18 E_DL_CipPhase 随本块
 *                         同文件发布；0.19 码位同行【级别】注释；0.20 验收向
 *                         量入头注释；R24 加药脉冲自清逻辑位于实例调用之后；
 *                         R25 bDone 单拍三律。
 * 红线自检 (Redline)    : R1 零全局变量表/外部变量引用 ✓｜R2 零物理 IO 地址 ✓
 *                         R3 纯 IEC 61131-3 ✓｜R4 越界/非有限值/互斥出口 ✓
 *                         R5 全变量中英双语同行注释 ✓｜R6 ENUM+CASE+ELSE ✓
 *                         R7 八实例主体最前部无条件刷新 ✓｜R8 全常量化 ✓
 *                         R24 TP/延时自清逻辑位于实例调用之后 ✓
 *                         R25 单拍标志生命周期三律 ✓
 * 设计要点 (Key notes)  : ① TACT 联锁暂停：温度/电导率/流量三路任一不达标
 *                           （下限 > 0 才校验）→ bPhaseHold、计时冻结、自动恢
 *                           复；暂停累计超 tHoldLimit → 相失败 0270（判失败
 *                           而非继续等）；TACT 信号非有限值按不达标保守侧暂
 *                           停（0172，不立即故障，防单点传感器抖动打断整批）；
 *                         ② 终冲洗特殊判据：以回液电导率 ≤ fRinseCondTarget
 *                           为完成条件（不以时间到为准），tRinseMax 兜底超时
 *                           → 0271；该相豁免零时长配方检查（偏离留档②）；
 *                         ③ 换相停泵间隔：相完成后先停泵 DL_CIP_SWITCH_PAUSE
 *                           再切阀（防混液，期间信息码 0173）；跳相仅由参数决
 *                           定——启动瞬间对启用数组做快照，运行中以快照推进
 *                           相序，中途改写启用数组视为「运行中跳相请求」一律
 *                           拒绝（信息码 0170，不生效）；
 *                         ④ 清洁许可：bCipComplete 仅全部启用相完成后置位；
 *                           中止即清除（中止即失去清洁许可）；复位路径清许可；
 *                           bOk = 完成保持态且全周期零偏差（以启动时偏差计数
 *                           快照比对）；
 *                         ⑤ 加药脉冲：电导率低于下限时每 DL_CIP_DOSING_PERIOD
 *                           一拍脉冲请求（R24 自清范式），非连续输出；
 *                         ⑥ 相位数组维度字面量 6（等同 DL_CIP_PHASE_MAX）与
 *                           常量同步维护（跨平台数组维度须编译期字面量）。
 * 偏离留档 (Deviation)  : 依 R11 头注释留档，共 2 条：
 *                         ① tCycle 增补引脚：相位计时累计需要时间基准，依公
 *                           约 0.10 增补（泳道 A 先例，公共约定强制项，非逐
 *                           组件条款）；
 *                         ② 零时长检查豁免终冲洗：规格「启用相目标时长为零 →
 *                           0272」未豁免任何相，但终冲洗以电导率判终点、时长
 *                           本就不参与其完成判据；按「终冲洗豁免 0272 检查」
 *                           实现。理由：终冲洗零时长在工艺上有意义（纯电导终
 *                           点）；影响：终冲洗配方时长域不校验。
 * 开源溯源 (Origin)     : 来源标签 cip-cleaning / isa-88-phase（RAW_NOTES_R8
 *                         S-10：CIP 原位清洗公开工程惯例——预冲/碱洗/中冲/酸
 *                         洗/终冲/消毒六相序、TACT 联锁暂停不计时、回液电导
 *                         率判终冲终点、回路就绪门控启泵、清洁状态（clean
 *                         status）放行生产、中止即失去许可（提取点①③④），
 *                         公开技术资料，仅借鉴相序分类与参数域；状态机、码
 *                         位、引脚契约 100% 本库独立设计，clean-room 未复制
 *                         源码。许可证说明：借鉴对象为公开技术惯例，无附带许
 *                         可限制；本文件为本库原创实现，随本库许可证发布）。
 * 验收向量 (Acceptance) :
 *   V1 六相全启用正常走完 → bCipComplete + bOk（零偏差）；
 *   V2 碱洗段温度低于下限 → 计时冻结 + bPhaseHold，恢复后继续；
 *   V3 暂停累计超 tHoldLimit → 0270 相失败锁存；
 *   V4 终冲洗回液电导降到终点 → 立即完成（不等 atPhaseTime）；
 *   V5 终冲洗超 tRinseMax → 0271；
 *   V6 abPhaseEnable[3]=FALSE → 跳过酸洗相（按启动快照）；
 *   V7 bAbort → 停泵排空 tDrainTime + bCipComplete=FALSE；
 *   V8 启用相 atPhaseTime=0 → 0272（终冲洗豁免，偏离留档②）。
 * 修订历史 (Revision)   :
 *   2026-11-15  v1.0.0  首版入库（Round 08 · DL_Process CIP 清洗件）
 *   2026-11-15  v1.0.1  R8 总监终审修复：终端态分支内的孤立空语句 `;`（非 IEC 61131-3 文法，statement_list 允许零条语句但不容纳孤立分号）改为纯注释占位分支，行为等价、跨平台可移植性合规。
 *============================================================================*)

(*-----------------------------------------------------------------------------
 * 枚举: E_DL_CipPhase（归属 FB_DL_CipCleaningSeq，与其同文件发布，公约 0.18）
 *----------------------------------------------------------------------------*)
TYPE E_DL_CipPhase :
(
    eIdle      := 0,   // 空闲：等启动 / Idle, awaiting start
    ePreRinse  := 10,  // 预冲洗（Pre-rinse）/ Pre-rinse phase
    eCaustic   := 20,  // 碱洗（Caustic wash）/ Caustic wash phase
    eIntRinse  := 30,  // 中间冲洗（Intermediate rinse）/ Intermediate rinse phase
    eAcid      := 40,  // 酸洗（Acid wash）/ Acid wash phase
    eFinalRinse:= 50,  // 终冲洗（Final rinse），电导率判终点 / Final rinse, conductivity end criterion
    eSanitize  := 60,  // 消毒（Sanitize）/ Sanitize phase
    eDone      := 70,  // 完成（bCipComplete），等复位 / Done, clean status granted
    eAbort     := 80,  // 中止：排空隔离，许可失效 / Aborted, drained and isolated, status revoked
    eFault     := 99   // 故障锁存 / Fault latched
) UINT;
END_TYPE

FUNCTION_BLOCK FB_DL_CipCleaningSeq
VAR_INPUT
    bEnable             : BOOL;             // 使能（Enable），FALSE=停泵停止加药（不主动排空），相位保持 / Enable, FALSE stops pumps and dosing, no drain
    bStart              : BOOL;             // 启动 CIP 周期（Start），上升沿受理（空闲/完成态）/ Start edge accepted at idle/done
    bAbort              : BOOL;             // 中止（Abort），电平最高优先 → 停泵 + 开排空 + 隔离 / Abort level, highest priority
    bReset              : BOOL;             // 复位（Reset），上升沿受理 / Rising edge resets fault and clean status
    bCircuitReady       : BOOL;             // 回路就绪（供货/回液阀位置确认），FALSE 禁止启泵与启动 / Circuit ready interlock
    abPhaseEnable       : ARRAY[0..5] OF BOOL;  // 各相启用（Phase enable）：0 预冲/1 碱/2 中冲/3 酸/4 终冲/5 消毒 / Phase enable flags, dim 6
    atPhaseTime         : ARRAY[0..5] OF TIME;  // 各相目标计时（Phase time），仅达标时段累计（终冲豁免，偏离留档②）/ Phase target durations
    afPhaseTempMin      : ARRAY[0..5] OF REAL;  // 各相温度下限（Temp min）[℃，0=不校验 / Phase temperature minimums, zero disables
    afPhaseCondMin      : ARRAY[0..5] OF REAL;  // 各相电导率下限（Conductivity min）[mS/cm，0=不校验 / Phase conductivity minimums, zero disables
    afPhaseFlowMin      : ARRAY[0..5] OF REAL;  // 各相流量下限（Flow min）[m³/h，0=不校验 / Phase flow minimums, zero disables
    fActTemp            : REAL;             // 实际温度（Actual temperature）[℃] / Actual temperature [degC]
    fActCond            : REAL;             // 实际电导率（Actual conductivity）[mS/cm]，供液或回液由调用方选择接点 / Actual conductivity [mS/cm]
    fActFlow            : REAL;             // 实际流量（Actual flow）[m³/h] / Actual flow [m3/h]
    fRinseCondTarget    : REAL := 0.1;      // 终冲洗回液电导率终点（Rinse conductivity target）[mS/cm] / Final-rinse conductivity end target
    tHoldLimit          : TIME := T#300S;   // 单相联锁暂停上限（Hold limit），超时判该相失败 / Per-phase hold limit, expiry = phase fail
    tRinseMax           : TIME := T#15M;    // 终冲洗最长延时（Rinse max time），电导未达标兜底上限 / Final-rinse maximum duration fallback
    tDrainTime          : TIME := T#60S;    // 中止后排空时长（Drain time）/ Abort drain duration
    tTempSetDelay       : TIME := T#0S;     // 升温/降温等待（Temp set delay），相开始先等待此窗不计时 / Temp settle delay before timing starts
    tCycle              : TIME := T#10MS;   // 任务扫描周期（Task cycle time）[ms]，由调用方按实际任务给，计时累计基准（偏离留档①）/ Task cycle time, timing base
END_VAR
VAR_OUTPUT
    ePhase              : E_DL_CipPhase := E_DL_CipPhase.eIdle; // 当前相位（Current phase）/ Current phase
    bBusy               : BOOL;             // 周期执行中（Busy），冲洗/消毒/换相/排空期 TRUE / TRUE during wash/sanitize/switch/drain
    bDone               : BOOL;             // 周期完成单拍（Done pulse），单拍生命周期三律 / One-scan completion pulse
    bOk                 : BOOL;             // 全相完成且无偏差（OK），完成保持态且零偏差 / OK verdict, done with zero deviations
    bPhaseHold          : BOOL;             // 相位暂停中（Phase hold），TACT 未达标计时冻结 / Phase hold, timing frozen
    bPhaseFail          : BOOL;             // 当前相失败（Phase fail），暂停超限锁存至复位 / Phase failed, latched until reset
    bCipComplete        : BOOL;             // CIP 完成许可（Clean status），供上层放行生产；中止/复位清除 / Clean status granted, revoked on abort/reset
    bCmdSupplyPump      : BOOL;             // 供液泵指令（Supply pump）/ Supply pump command
    bCmdReturnPump      : BOOL;             // 回液泵指令（Return pump）/ Return pump command
    bCmdDosing          : BOOL;             // 加药泵指令（Dosing pump），电导率低于下限时脉冲式请求 / Dosing pulse request
    bCmdHeat            : BOOL;             // 加热（蒸汽阀）指令（Heat）/ Heat command
    bCmdDrain           : BOOL;             // 排空阀指令（Drain valve），中止排空期 / Drain valve command
    fTempSetpoint       : REAL;             // 温度设定（Temp setpoint）[℃]，取当前相下限 + 2.0 ℃ 裕量（工艺经验值）/ Temp setpoint, phase min plus margin
    tPhaseElapsed       : TIME := T#0S;     // 当前相已累计计时（Phase elapsed），仅达标时段 / Accumulated phase time, qualified periods only
    nDeviationCount     : UDINT;            // 偏差计数（Deviation counter），每次暂停/失败 +1，供审计 / Deviation counter for audit
    bError              : BOOL;             // 故障锁存（Error），仅故障级码 / Latched error, fault codes only
    uErrorId            : UDINT;            // 故障码（Error code），16#0005_xxxx 段，0=无故障 / Error code, fault-level priority
END_VAR
VAR
    _ePhase             : E_DL_CipPhase := E_DL_CipPhase.eIdle;   // 内部相位（Internal phase）/ Internal phase
    _nPhaseIdx          : UINT := UINT#6;   // 当前相索引（Current phase index）[-]，0..5；6=哨兵（无活动相）/ Index 0..5, 6 = sentinel none
    _nNextIdx           : UINT;             // 下一相索引（Next phase index）[-]，哨兵 6 / Next phase index, sentinel 6
    _bEnterPhase        : BOOL;             // 进入相位单拍（Enter phase one-shot），索引→枚举映射触发 / Phase-entry one-shot for mapping
    _bPhaseActive       : BOOL;             // 相位执行中派生（Phase active derived）/ Wash phase active derived
    _bFaultLatch        : BOOL;             // 故障锁存标志（Fault latch flag），仅复位路径清除 / Fault latch, cleared only via reset path
    _uErrorIdInt        : UDINT;            // 内部故障级码寄存（Internal fault-level register）/ Internal fault-level register
    _uInfoCode          : UDINT;            // 本拍信息级码（Info code this cycle），瞬时型每拍重算 / Transient info code
    _bSwitchPause       : BOOL;             // 换相停泵间隔（Switch pause），防混液 / Switch pause between phases
    _tPhaseElapsedInt   : TIME := T#0S;     // 内部相位计时（Internal phase elapsed）/ Internal phase elapsed
    _bTempHold          : BOOL;             // 温度联锁暂停（Temperature hold）/ Temperature interlock hold
    _bCondHold          : BOOL;             // 电导率联锁暂停（Conductivity hold）/ Conductivity interlock hold
    _bFlowHold          : BOOL;             // 流量联锁暂停（Flow hold）/ Flow interlock hold
    _bHold              : BOOL;             // 联锁暂停归并（Hold merged）/ Merged hold flag
    _bHoldPrev          : BOOL;             // 上拍暂停态（Hold previous scan），进入沿计数用 / Hold previous scan, entry edge
    _bDosePulse         : BOOL;             // 加药脉冲单拍（Dosing pulse one-shot）/ Dosing pulse one-shot
    _bPhaseDone         : BOOL;             // 当前相完成（Phase done）/ Current phase completed
    _bDrainDone         : BOOL;             // 排空完成（Drain done）/ Drain completed
    _bParamEdited       : BOOL;             // 启用数组中途改写（Enable array edited mid-run），跳相拒绝判据 / Enable array edited mid-run
    _nIdx               : UINT;             // 循环索引（Loop index）[-] / Loop index
    _fTempMin           : REAL;             // 当前相温度下限（Phase temp minimum）[℃] / Current phase temperature minimum
    _fCondMin           : REAL;             // 当前相电导率下限（Phase cond minimum）[mS/cm] / Current phase conductivity minimum
    _fFlowMin           : REAL;             // 当前相流量下限（Phase flow minimum）[m³/h] / Current phase flow minimum
    _bFiniteTact        : BOOL;             // 三路 TACT 信号有限归并（TACT finite merged）/ Merged TACT finite verdict
    _abEnableSnap       : ARRAY[0..5] OF BOOL;  // 启用数组启动快照（Enable snapshot at start），运行中改写不生效 / Enable snapshot taken at start
    _nDevStart          : UDINT;            // 启动时偏差计数快照（Deviation snapshot at start），零偏差判定基准 / Deviation count snapshot at start
    _fbTrigStart        : R_TRIG;           // 启动沿（Start edge detector）/ Start edge detector
    _fbTrigReset        : R_TRIG;           // 复位沿（Reset edge detector）/ Reset edge detector
    _fbTonHold          : TON;              // 联锁暂停上限（Hold limit timer）/ Hold limit timer
    _fbTonDose          : TON;              // 加药脉冲周期（Dosing period timer）/ Dosing period timer
    _fbTonSwitch        : TON;              // 换相停泵间隔（Switch pause timer）/ Switch pause timer
    _fbTonDrain         : TON;              // 排空时长（Drain duration timer）/ Drain duration timer
    _fbTonTempDelay     : TON;              // 升降温等待窗（Temp settle delay timer）/ Temp settle delay timer
    _fbTonRinseMax      : TON;              // 终冲洗最长延时（Rinse max timer）/ Final-rinse max timer
END_VAR
VAR CONSTANT
    DL_CIP_PHASE_MAX    : UINT := 6;        // 相位数上限（Max phases）[-]，与数组维度字面量 6 同步 / Phase count, sync with literal dim 6
    DL_CIP_IDX_NONE     : UINT := 6;        // 无活动相哨兵索引（Sentinel index for none）[-] / Sentinel index, none active
    DL_CIP_IDX_FINAL    : UINT := 4;        // 终冲洗相索引（Final-rinse index）[-] / Final-rinse phase index
    DL_CIP_REAL_MAX     : REAL := 3.4E38;   // 单精度有限值判据幅值（Finite magnitude bound）/ Finite magnitude bound for REAL inputs
    DL_CIP_TEMP_MARGIN  : REAL := 2.0;      // 温度设定裕量（Temp setpoint margin）[℃]，工艺经验值 / Temperature margin, process experience
    DL_CIP_DOSING_PERIOD: TIME := T#5S;     // 加药脉冲周期（Dosing pulse period）/ Dosing pulse period
    DL_CIP_SWITCH_PAUSE : TIME := T#2S;     // 换相停泵间隔（Switch pause duration），防混液 / Pump-off pause between phases
    DL_CIP_ERR_HOLD     : UDINT := 16#0005_0270; // 0005_0270 单相联锁暂停超限（相失败）【故障级】/ Phase hold limit exceeded, fault level
    DL_CIP_ERR_RINSE    : UDINT := 16#0005_0271; // 0005_0271 终冲洗超最长延时未达电导终点【故障级】/ Final rinse over max duration, fault level
    DL_CIP_ERR_ZEROTIME : UDINT := 16#0005_0272; // 0005_0272 启用相目标时长为零【故障级】/ Enabled phase with zero duration, fault level
    DL_CIP_ERR_NOREADY  : UDINT := 16#0005_0273; // 0005_0273 回路未就绪强行启动【故障级】/ Started with circuit not ready, fault level
    DL_CIP_ERR_STATE    : UDINT := 16#0005_0274; // 0005_0274 非法状态兜底【故障级】/ Illegal state fallback, fault level
    DL_CIP_INFO_SKIP    : UDINT := 16#0005_0170; // 0005_0170 运行中跳相请求被拒（启用数组中途改写不生效）【信息级】/ Mid-run phase skip refused, info level
    DL_CIP_INFO_NOREADY : UDINT := 16#0005_0171; // 0005_0171 回路未就绪，泵指令被抑制【信息级】/ Pump suppressed, circuit not ready, info level
    DL_CIP_INFO_NAN     : UDINT := 16#0005_0172; // 0005_0172 TACT 信号非有限值，保守侧暂停【信息级】/ TACT non-finite, conservative hold, info level
    DL_CIP_INFO_SWITCH  : UDINT := 16#0005_0173; // 0005_0173 相切换停泵间隔中【信息级】/ Pump-off switch pause, info level
END_VAR

// ============================================================================
// 段 1｜实例无条件周期刷新（R7/0.5：严禁置于 IF/CASE 分支内）
//      Unconditional per-cycle refresh of all instances (R7/0.5)
// ============================================================================
_fbTrigStart(CLK := bStart);            // 启动沿（Start edge）
_fbTrigReset(CLK := bReset);            // 复位沿（Reset edge）

// 相位执行中派生（Phase active derived）
_bPhaseActive := (_ePhase = E_DL_CipPhase.ePreRinse) OR (_ePhase = E_DL_CipPhase.eCaustic)
              OR (_ePhase = E_DL_CipPhase.eIntRinse) OR (_ePhase = E_DL_CipPhase.eAcid)
              OR (_ePhase = E_DL_CipPhase.eFinalRinse) OR (_ePhase = E_DL_CipPhase.eSanitize);

// 联锁暂停上限（仅执行相计时，暂停解除/相失败自动断输入归零）
// Hold limit timer (armed in active phases, auto reset on release)
_fbTonHold(IN := _bPhaseActive AND bEnable AND _bHold AND (NOT _bSwitchPause), PT := tHoldLimit);
// 加药脉冲周期（仅电导暂停期计时；R24：脉冲自清逻辑在段 3 实例调用之后）
// Dosing period timer (armed on conductivity hold; R24 self-clear after call)
_fbTonDose(IN := _bCondHold AND bEnable AND (NOT _bDosePulse) AND (NOT _bSwitchPause), PT := DL_CIP_DOSING_PERIOD);
// 换相停泵间隔（Switch pause timer）
_fbTonSwitch(IN := _bSwitchPause, PT := DL_CIP_SWITCH_PAUSE);
// 排空时长（仅中止相且未排空完成时计时 / Drain timer, abort phase until done）
_fbTonDrain(IN := (_ePhase = E_DL_CipPhase.eAbort) AND (NOT _bDrainDone), PT := tDrainTime);
// 升降温等待窗（相开始后到窗才允许计时 / Temp settle delay before timing allowed）
_fbTonTempDelay(IN := _bPhaseActive AND bEnable AND (NOT _bSwitchPause), PT := tTempSetDelay);
// 终冲洗最长延时（Final-rinse max timer）
_fbTonRinseMax(IN := (_ePhase = E_DL_CipPhase.eFinalRinse) AND bEnable, PT := tRinseMax);

// ============================================================================
// 段 2｜信息级预清零 + 输出默认赋值（0.9：任何早退路径输出确定）
//      Info preset + output defaults
// ============================================================================
_uInfoCode := 0;                        // 信息级瞬时型每拍重算（Transient info recomputed each scan）
bDone := FALSE;                         // 完成单拍先清零（R25：置位-消费-复位同周期闭环）/ Done pulse preset FALSE (R25)
bCmdSupplyPump := FALSE;                // 泵/阀/加药/加热指令默认安全侧全关（Commands preset closed）
bCmdReturnPump := FALSE;
bCmdDosing := FALSE;
bCmdHeat := FALSE;
bCmdDrain := FALSE;
fTempSetpoint := 0.0;                   // 温度设定默认零（Temp setpoint default zero）
bPhaseHold := FALSE;                    // 暂停/失败/判定默认清（Hold, fail, verdict preset）
bPhaseFail := FALSE;
bOk := FALSE;

// 当前相参数取值（索引先判域，防越界）
// Current phase parameter fetch (index bounded first)
IF _nPhaseIdx < DL_CIP_PHASE_MAX THEN
    _fTempMin := afPhaseTempMin[_nPhaseIdx];   // 当前相温度下限（Phase temp minimum）
    _fCondMin := afPhaseCondMin[_nPhaseIdx];   // 当前相电导率下限（Phase cond minimum）
    _fFlowMin := afPhaseFlowMin[_nPhaseIdx];   // 当前相流量下限（Phase flow minimum）
ELSE
    _fTempMin := 0.0;                   // 越界防御默认（Bounded default）
    _fCondMin := 0.0;
    _fFlowMin := 0.0;
END_IF

// TACT 信号非有限值防御（自比等价式，归并三路）
// TACT non-finite defense (self-comparison equivalence, merged)
_bFiniteTact := (fActTemp >= (-DL_CIP_REAL_MAX)) AND (fActTemp <= DL_CIP_REAL_MAX)
           AND (fActCond >= (-DL_CIP_REAL_MAX)) AND (fActCond <= DL_CIP_REAL_MAX)
           AND (fActFlow >= (-DL_CIP_REAL_MAX)) AND (fActFlow <= DL_CIP_REAL_MAX);

// ============================================================================
// 段 3｜TACT 联锁判定与计时累计（仅执行相；R24 脉冲自清在实例调用之后）
//      TACT interlock and timing accumulation (R24 pulse self-clear after call)
// ============================================================================
IF _bPhaseActive AND bEnable AND (NOT _bSwitchPause) THEN
    _bTempHold := (_fTempMin > 0.0) AND ((NOT _bFiniteTact) OR (fActTemp < _fTempMin));
    _bCondHold := (_fCondMin > 0.0) AND ((NOT _bFiniteTact) OR (fActCond < _fCondMin));
    _bFlowHold := (_fFlowMin > 0.0) AND ((NOT _bFiniteTact) OR (fActFlow < _fFlowMin));
    _bHold := _bTempHold OR _bCondHold OR _bFlowHold;   // 三路归并（Merged hold）
    IF (NOT _bFiniteTact) AND _bHold THEN
        _uInfoCode := DL_CIP_INFO_NAN;   // 0005_0172 TACT 非有限值保守侧暂停【信息级】/ TACT non-finite, info level
    END_IF
    // 暂停进入沿：偏差计数 +1（Hold entry edge: deviation count increment）
    IF _bHold AND (NOT _bHoldPrev) THEN
        nDeviationCount := nDeviationCount + UINT#1;
    END_IF
    // 计时累计：联锁全达标且升降温等待窗已过（Timing: interlocks met and delay elapsed）
    IF (NOT _bHold) AND _fbTonTempDelay.Q THEN
        _tPhaseElapsedInt := _tPhaseElapsedInt + tCycle;
        tPhaseElapsed := _tPhaseElapsedInt;              // 出口计时同步（Outlet elapsed sync）
    END_IF
ELSE
    _bTempHold := FALSE;                // 非执行相暂停清零（Hold cleared off-phase）
    _bCondHold := FALSE;
    _bFlowHold := FALSE;
    _bHold := FALSE;
END_IF
_bHoldPrev := _bHold;                   // 登记本拍暂停态供下拍沿判定（Register hold for edge）

// R24 范式：加药脉冲单拍自清（实例调用之后置位，下一拍 IN 断自动复位）
// R24 pattern: dosing pulse set after instance call, auto-resets next scan
_bDosePulse := _fbTonDose.Q;            // 脉冲单拍登记（Pulse one-shot registered）

// 相失败监视：暂停累计超上限（Phase fail monitor: hold limit exceeded）
IF _fbTonHold.Q AND (NOT _bFaultLatch) THEN
    _bFaultLatch := TRUE;               // 相失败锁存（Phase fail latch）
    _uErrorIdInt := DL_CIP_ERR_HOLD;    // 0005_0270 单相联锁暂停超限【故障级】/ Phase hold exceeded, fault level
    _ePhase := E_DL_CipPhase.eFault;
END_IF

// 终冲洗兜底监视：超最长延时未达电导终点（Final-rinse max monitor）
IF _fbTonRinseMax.Q AND (NOT _bFaultLatch) THEN
    _bFaultLatch := TRUE;               // 终冲超时锁存（Final-rinse timeout latch）
    _uErrorIdInt := DL_CIP_ERR_RINSE;   // 0005_0271 终冲洗超最长延时【故障级】/ Final-rinse timeout, fault level
    _ePhase := E_DL_CipPhase.eFault;
END_IF

// ============================================================================
// 段 4｜核心相位状态机（ENUM + CASE，含 ELSE 非法状态兜底）
//      Core phase state machine (ENUM + CASE with ELSE fallback)
// ============================================================================
IF bEnable AND (NOT _bFaultLatch) THEN
    IF bAbort AND (_ePhase <> E_DL_CipPhase.eIdle) AND (_ePhase <> E_DL_CipPhase.eAbort) THEN
        // 中止电平拦截：排空隔离、清洁许可失效（Abort intercept: drain, status revoked）
        bCipComplete := FALSE;          // 中止即失去清洁许可（Clean status revoked on abort）
        _bDrainDone := FALSE;           // 排空重新武装（Drain re-armed）
        _ePhase := E_DL_CipPhase.eAbort;
    ELSE
        CASE _ePhase OF

            E_DL_CipPhase.eIdle: // 空闲：等启动沿
                IF _fbTrigStart.Q THEN
                    IF NOT bCircuitReady THEN
                        _bFaultLatch := TRUE;                // 回路未就绪强行启动（Started not ready）
                        _uErrorIdInt := DL_CIP_ERR_NOREADY;  // 0005_0273 回路未就绪启动【故障级】/ Started not ready, fault level
                        _ePhase := E_DL_CipPhase.eFault;
                    ELSE
                        // 启动前配方检查：启用相零时长（终冲豁免，偏离留档②）
                        // Pre-start recipe check: enabled zero-duration (final rinse exempt)
                        FOR _nIdx := UINT#0 TO DL_CIP_PHASE_MAX - UINT#1 DO
                            IF abPhaseEnable[_nIdx] AND (atPhaseTime[_nIdx] = T#0MS)
                            AND (_nIdx <> DL_CIP_IDX_FINAL) THEN
                                _bFaultLatch := TRUE;                 // 零时长相锁存（Zero duration latch）
                                _uErrorIdInt := DL_CIP_ERR_ZEROTIME;  // 0005_0272 启用相零时长【故障级】/ Zero duration, fault level
                            END_IF
                        END_FOR
                        IF NOT _bFaultLatch THEN
                            // 启用数组快照 + 偏差基准快照（Snapshot enable array and deviation base）
                            FOR _nIdx := UINT#0 TO DL_CIP_PHASE_MAX - UINT#1 DO
                                _abEnableSnap[_nIdx] := abPhaseEnable[_nIdx];
                            END_FOR
                            _nDevStart := nDeviationCount;
                            // 找首个启用相进入（Find first enabled phase）
                            _nPhaseIdx := DL_CIP_IDX_NONE;            // 哨兵：无启用相（Sentinel: none enabled）
                            FOR _nIdx := UINT#0 TO DL_CIP_PHASE_MAX - UINT#1 DO
                                IF (_nPhaseIdx = DL_CIP_IDX_NONE) AND _abEnableSnap[_nIdx] THEN
                                    _nPhaseIdx := _nIdx;              // 首个启用相（First enabled phase）
                                END_IF
                            END_FOR
                            IF _nPhaseIdx < DL_CIP_PHASE_MAX THEN
                                _tPhaseElapsedInt := T#0S;            // 相计时清零（Phase elapsed reset）
                                tPhaseElapsed := T#0S;
                                _bSwitchPause := FALSE;
                                _bPhaseDone := FALSE;
                                _bEnterPhase := TRUE;                 // 触发索引→枚举映射（Arm phase mapping）
                            ELSE
                                _ePhase := E_DL_CipPhase.eDone;       // 全相禁用直接完成（All disabled, straight done）
                                bCipComplete := TRUE;                 // 清洁许可（Clean status granted）
                                bDone := TRUE;                        // 完成单拍（R25 本拍闭环）/ Done pulse (R25)
                            END_IF
                        END_IF
                    END_IF
                END_IF

            E_DL_CipPhase.ePreRinse, E_DL_CipPhase.eCaustic, E_DL_CipPhase.eIntRinse,
            E_DL_CipPhase.eAcid, E_DL_CipPhase.eFinalRinse, E_DL_CipPhase.eSanitize:
                // 六相公共执行分支（Common wash-phase branch）
                IF (_nPhaseIdx < DL_CIP_PHASE_MAX) AND (NOT _bSwitchPause) THEN
                    // 终冲洗特殊判据：回液电导率 ≤ 终点即完成（不以时间到为准）
                    // Final rinse: conductivity end criterion (time not decisive)
                    IF (_ePhase = E_DL_CipPhase.eFinalRinse) AND _bFiniteTact
                    AND (fActCond <= fRinseCondTarget) AND (NOT _bHold) THEN
                        _bPhaseDone := TRUE;              // 电导终点达成（Conductivity end met）
                    ELSIF (_ePhase <> E_DL_CipPhase.eFinalRinse)
                    AND (_tPhaseElapsedInt >= atPhaseTime[_nPhaseIdx]) THEN
                        _bPhaseDone := TRUE;              // 目标时长达成（Target duration met）
                    END_IF
                    IF _bPhaseDone THEN
                        _bSwitchPause := TRUE;            // 相完成进入停泵间隔（Phase done, pump-off pause）
                        _uInfoCode := DL_CIP_INFO_SWITCH; // 0005_0173 换相停泵间隔【信息级】/ Switch pause, info level
                    END_IF
                END_IF

            E_DL_CipPhase.eDone: // 完成保持：等复位（复位路径在段 6）
                // 等复位（Awaiting reset）

            E_DL_CipPhase.eAbort: // 中止排空：排空时长到后保持等待复位
                IF _fbTonDrain.Q THEN
                    _bDrainDone := TRUE;              // 排空完成（Drain completed）
                END_IF

            E_DL_CipPhase.eFault: // 故障锁存：等复位
                // 等复位（Awaiting reset）

            ELSE // 非法状态兜底（本块专用码位）
                _bFaultLatch := TRUE;
                _uErrorIdInt := DL_CIP_ERR_STATE;     // 0005_0274 非法状态兜底【故障级】/ Illegal state fallback, fault level
                _ePhase := E_DL_CipPhase.eFault;
        END_CASE
    END_IF
END_IF

// ============================================================================
// 段 5｜换相推进 + 索引→枚举映射 + 运行中改写检测（索引先判域）
//      Phase advance, index-to-enum mapping, mid-run edit detection (bounded)
// ============================================================================
IF _bSwitchPause AND _fbTonSwitch.Q AND (NOT _bFaultLatch) THEN
    _bSwitchPause := FALSE;             // 停泵间隔结束（Pause finished）
    _bPhaseDone := FALSE;
    // 从当前相之后按启动快照找下一启用相（Next enabled phase after current, snapshot-based）
    _nNextIdx := DL_CIP_IDX_NONE;       // 哨兵：无后续启用相（Sentinel: none left）
    IF _nPhaseIdx + UINT#1 <= DL_CIP_PHASE_MAX - UINT#1 THEN
        FOR _nIdx := _nPhaseIdx + UINT#1 TO DL_CIP_PHASE_MAX - UINT#1 DO
            IF (_nNextIdx = DL_CIP_IDX_NONE) AND _abEnableSnap[_nIdx] THEN
                _nNextIdx := _nIdx;     // 下一启用相（Next enabled phase）
            END_IF
        END_FOR
    END_IF
    IF _nNextIdx < DL_CIP_PHASE_MAX THEN
        _nPhaseIdx := _nNextIdx;        // 推进到下一相（Advance to next phase）
        _tPhaseElapsedInt := T#0S;      // 相计时清零（Phase elapsed reset）
        tPhaseElapsed := T#0S;
        _bEnterPhase := TRUE;           // 触发索引→枚举映射（Arm phase mapping）
    ELSE
        _ePhase := E_DL_CipPhase.eDone; // 全部启用相完成（All enabled phases done）
        bCipComplete := TRUE;           // 清洁许可（Clean status granted）
        bDone := TRUE;                  // 完成单拍（R25 本拍闭环）/ Done pulse (R25)
    END_IF
END_IF

// 相位索引→枚举映射（进入相单拍执行；越界防御）
// Index-to-enum mapping (on phase-entry one-shot, bounded)
IF _bEnterPhase AND (_nPhaseIdx < DL_CIP_PHASE_MAX) THEN
    CASE _nPhaseIdx OF
        UINT#0: _ePhase := E_DL_CipPhase.ePreRinse;    // 预冲洗（Pre-rinse）
        UINT#1: _ePhase := E_DL_CipPhase.eCaustic;     // 碱洗（Caustic）
        UINT#2: _ePhase := E_DL_CipPhase.eIntRinse;    // 中间冲洗（Intermediate）
        UINT#3: _ePhase := E_DL_CipPhase.eAcid;        // 酸洗（Acid）
        UINT#4: _ePhase := E_DL_CipPhase.eFinalRinse;  // 终冲洗（Final rinse）
        UINT#5: _ePhase := E_DL_CipPhase.eSanitize;    // 消毒（Sanitize）
        ELSE _ePhase := E_DL_CipPhase.eIdle;           // 防御回空闲（Bounded default）
    END_CASE
    _bEnterPhase := FALSE;              // 映射消费（Mapping consumed）
END_IF

// 运行中启用数组改写检测：视为跳相请求一律拒绝（不生效，仅信息码 0170）
// Mid-run enable edit detection: treated as skip request, refused (info 0170)
IF _bPhaseActive THEN
    _bParamEdited := FALSE;             // 改写判据预清（Edit flag preset）
    FOR _nIdx := UINT#0 TO DL_CIP_PHASE_MAX - UINT#1 DO
        IF abPhaseEnable[_nIdx] <> _abEnableSnap[_nIdx] THEN
            _bParamEdited := TRUE;      // 检测到改写（Edit detected）
        END_IF
    END_FOR
    IF _bParamEdited THEN
        _uInfoCode := DL_CIP_INFO_SKIP; // 0005_0170 运行中跳相请求被拒【信息级】/ Mid-run skip refused, info level
    END_IF
END_IF

// ============================================================================
// 段 6｜复位路径 + 输出派生（R15：故障/许可仅复位路径清；0171 泵抑制）
//      Reset path + outlet derivation (R15; pump suppression on not-ready)
// ============================================================================
IF _fbTrigReset.Q THEN
    _bFaultLatch := FALSE;              // 故障锁存解除（Fault latch released）
    _uErrorIdInt := 16#0000_0000;       // 故障码清零（Fault code cleared）
    bCipComplete := FALSE;              // 清洁许可随复位清除（Clean status cleared on reset）
    _bDrainDone := FALSE;               // 排空标志复位（Drain flag reset）
    _nPhaseIdx := DL_CIP_IDX_NONE;      // 相索引回哨兵（Index back to sentinel）
    IF (_ePhase = E_DL_CipPhase.eFault) OR (_ePhase = E_DL_CipPhase.eAbort)
    OR (_ePhase = E_DL_CipPhase.eDone) THEN
        _ePhase := E_DL_CipPhase.eIdle; // 终态回空闲（Terminal phases back to idle）
        _tPhaseElapsedInt := T#0S;
        tPhaseElapsed := T#0S;
    END_IF
END_IF

// 相失败出口：仅联锁暂停超限锁存为相失败，锁存至复位（与 bPhaseHold 不同真）
// Phase fail outlet: hold-limit latch only, held until reset (exclusive with hold)
IF _bFaultLatch AND (_uErrorIdInt = DL_CIP_ERR_HOLD) THEN
    bPhaseFail := TRUE;                 // 相失败锁存出口（Phase fail latched outlet）
END_IF

// 泵/加药/加热指令：执行相且回路就绪且非停泵间隔且无故障（0171 泵抑制每拍重算）
// Pump/dosing/heat: active phase AND circuit ready AND not in pause AND no fault
IF _bPhaseActive AND bEnable AND bCircuitReady AND (NOT _bSwitchPause) AND (NOT _bFaultLatch) THEN
    bCmdSupplyPump := TRUE;             // 供液泵开（Supply pump on）
    bCmdReturnPump := TRUE;             // 回液泵开（Return pump on）
    bCmdHeat := _bTempHold;             // 加热：温度暂停期（Heat on temperature hold）
    bCmdDosing := _bDosePulse;          // 加药：电导暂停脉冲（Dosing pulse on cond hold）
END_IF
IF _bPhaseActive AND bEnable AND (NOT bCircuitReady) AND (NOT _bFaultLatch) THEN
    _uInfoCode := DL_CIP_INFO_NOREADY;  // 0005_0171 回路未就绪泵被抑制【信息级】/ Pump suppressed, info level
END_IF

// 排空阀：中止相排空期内（Drain valve during abort drain window）
bCmdDrain := (_ePhase = E_DL_CipPhase.eAbort) AND (NOT _bDrainDone);

// 温度设定：当前相下限 + 裕量（下限 0=不校验则设定 0）
// Temp setpoint: phase minimum plus margin (zero minimum = zero setpoint)
IF _bPhaseActive AND (_fTempMin > 0.0) THEN
    fTempSetpoint := _fTempMin + DL_CIP_TEMP_MARGIN;   // 抬高 2 ℃ 裕量（Margin applied）
END_IF

// 判定出口：完成保持态且全周期零偏差（以启动偏差快照比对）
// Verdict outlet: done hold with zero whole-cycle deviations (vs start snapshot)
IF _ePhase = E_DL_CipPhase.eDone THEN
    bOk := (nDeviationCount = _nDevStart);   // 零偏差判定（Zero-deviation verdict）
END_IF

bBusy := _bPhaseActive OR (_ePhase = E_DL_CipPhase.eAbort);   // 执行中派生（Busy derived）

ePhase := _ePhase;                       // 相位镜像（Phase mirror）

// ============================================================================
// 段 7｜bError/uErrorId 出口（R21：bError 显式排除信息级码）
//      Outlets: bError excludes info codes (R21)
// ============================================================================
bError := _bFaultLatch;                  // 故障级派生式（Fault-level derived form）
IF _bFaultLatch THEN
    uErrorId := _uErrorIdInt;            // 故障级码优先透出（Fault-level priority）
ELSE
    uErrorId := _uInfoCode;              // 无故障时透出本拍信息级码（Transient info code）
END_IF
END_FUNCTION_BLOCK

(* ---- FB_DL_CompressorSurgeGuard.st ---- *)
(*==============================================================================
 * 组件名称 (Component)  : FB_DL_CompressorSurgeGuard
 * 溯源说明 (Provenance): 道莅 clean-room 防御性实现（IEC 61131-3 纯净实现，闭源文档仅借语义，零代码行）
 * 所属子库 (Sublibrary) : DL_Process / ProcessSafety
 * 当前版本 (Version)    : 1.0.0
 * 兼容性   (Platform)   : CODESYS 3.5 / TwinCAT 3 / 汇川 InoProShop / 施耐德
 *                         Machine Expert；纯 IEC 61131-3（第 3 版），仅用
 *                         Standard.library 的 TON / LIMIT / MAX / ABS 与
 *                         子库内 FB_DL_RateLimiter（DL_Algo，Level 1）
 * 组件分类 (Category)   : 功能块（FUNCTION_BLOCK）· 压缩机防喘振
 * 功能一句话 (Summary)  : 按压比修正最小流量危险线，流量跌破危险线持续确认后
 *                         快开放空阀，流量回升并越出回差带后慢关，全程给出
 *                         压比、喘振风险与放空动作可观测位。
 *
 * 本件存在的意义 (Why this unit exists)
 *   喘振是压缩机的爆炸级失效模式：流量低于临界值时机组进入周期性倒流振荡，
 *   十几秒内即可损坏转子与密封。库内没有任何件管这条保护律。本件把
 *   「最小流量线按压比修正 + 确认延时 + 快开慢关 + 回差恢复」四件事写成一件，
 *   且只编排已收口能力（斜率先行由 FB_DL_RateLimiter 承担，不复制其算法）。
 *
 * 危险线口径 (Danger line)
 *   fFlowDanger = fFlowMinLine × (1 + fSurgeMargin × (压比 − 1))
 *   线性近似：压比越高，同样流量下越接近喘振，故危险线上抬。公式与系数
 *   100 % 自有，不引用任何厂商曲线。压比夹到 ≥ 1.0——压比小于 1 的测量值
 *   不可信（吸入压力大于排出压力），若直接代入会让危险线低于最小流量线，
 *   保护范围凭空缩小，故按 1.0 处理并留档。
 *
 * 两条安全方向相反的规则（并列写死，不得只做其一）
 *   ① 参数非法（最小流量线/裕度/斜率为非正、吸入压力 ≤ 0）→ 故障 030B、
 *      阀**全开**：宁可放空不可喘振（放空只浪费能量，喘振会毁机）；
 *   ② 任一输入非有限 → 故障 030C、**保持末次阀位**：坏值不得成为关阀理由
 *      （P0 级，与①方向相反，两条都必须写死，见段 9）。
 *
 * 边界安全 (Boundary)
 *   - 流量低于危险线持续 tConfirm → eRiskBlowoff，阀按 fOpenRamp 快开；
 *   - 流量恢复到 fFlowDanger ×(1 + DL_SURGE_HYST) 以上 → eRecovering，
 *     阀按 fCloseRamp 慢关；**关到 0 才回 eNormal**——eRiskBlowoff 不得被
 *     eNormal 直接抢占（R41 回差家族），也不存在「风险刚解除就全关」的路径；
 *   - 失能 → 阀仍按 fCloseRamp 关闭（不阶跃），bBlowoffActive := FALSE，
 *     bSurgeRisk 保持可观测（停机期间仍要让 HMI 看到风险）；
 *   - CASE 落 ELSE 置 030D 并回 eFault；本件无复位引脚，故障态在原因消失后
 *     自动回 eNormal（无台账需保持，与安全阀台账件语义不同，已留档）；
 *   - 斜坡组合调用按 R36 处理**首次扫描退出跟踪的首拍**：阀位经
 *     FB_DL_RateLimiter 跟踪注入（bTrack / fTrackValue）而非直接赋值，
 *     首拍与「非有限保持 → 恢复」首拍都不产生阶跃。
 * 依赖与码位纪律
 *   子件 FB_DL_RateLimiter 的错误码属 16#0002_ 段（DL_Algo 属主），
 *   **不并入**本件码位体系（R70② 段属主唯一）；本件参数闸门已把斜率钳成
 *   有限正值、采样周期恒 ≥ 下限，故子件两条错误路径结构性不可达。
 *
 * 错误码    : 16#0005_01DA 流量低于危险线，放空阀已打开——信息级，保护动作
 *             16#0005_01DB 流量已回升越出回差带，退出放空——信息级，恢复动作
 *             16#0005_030B 防喘振参数非法（含吸入压力 ≤ 0），阀全开——故障级
 *             16#0005_030C 输入非有限，保持末次阀位——故障级，坏值不得关阀
 *             16#0005_030D 状态机落 ELSE 兜底（非法状态）——故障级，回 eFault
 * 码位总账  : 16#0005_01DA 用 / 16#0005_01DB 用 ｜ 16#0005_030B 用 / 16#0005_030C 用 / 16#0005_030D 用
 * 状态机    : E_DL_SurgeState（eIdle / eNormal / eRiskBlowoff / eRecovering / eFault），
 *             CASE 含 ELSE 兜底，ELSE 置 16#0005_030D 并回 eFault；失能无条件回 eIdle
 * 采样约定  : 每任务周期调用一次；斜率 [%/s] 依赖 tSample 引脚（禁读系统时钟）
 * 依赖说明  : DL_Process 可依赖 Level 0/1，本件只**组合调用** FB_DL_RateLimiter，
 *             不复制其斜坡算法（R36 手算首拍跟踪见上）
 * 验收向量  : V1 吸入 100 / 排出 300 / 流量 2000 / 最小线 500 / 裕度 0.10
 *               → 压比 3.0，危险线 500×(1+0.10×2)=600，流量高于危险线 → eNormal，
 *                 阀 0%，bSurgeRisk = FALSE
 *             V2 流量跌到 500（< 600）持续 200 ms → eRiskBlowoff，阀按 20 %/s 快开，
 *                 eErr = 01DA，bBlowoffActive = TRUE
 *             V3 V2 后流量回到 700（> 600×1.15=690）→ eRecovering，阀按 1 %/s 慢关，
 *                 eErr = 01DB；关到 0 才回 eNormal（回差主向量）
 *             V4 fFlowMinLine = 0 → 阀 100 %，eErr = 030B，bError = TRUE
 *             V5 fDischargePress = NaN → 阀保持末次值，eErr = 030C（保持主向量）
 *             V6 fSuctionPress = 0 → 按参数类 030B，阀全开（压比无意义主向量）
 *             V7 bEnable = FALSE → 阀按 1 %/s 降到 0，bBlowoffActive = FALSE，
 *                bSurgeRisk 仍随流量可观测
 * 红线自检  : 全局变量声明零使用 / 外部变量访问零使用 / 物理地址零使用 ｜ 纯 IEC 61131-3 ｜ 压比除零
 *             前置闸（吸入压力 > 0 才做除法）｜ 浮点只用大小与容差比较 ｜ 无循环
 *             ｜ 全变量双语同行注释 ｜ ENUM + CASE 含 ELSE ｜ TON 在主体最前部
 *             无条件刷新 ｜ 斜率/回差全部常量化，无魔法数
 * 修订历史  : 2026-11-16  v1.0.0  首版入库（R22 · 批 2 · 过程单元保护）
 *============================================================================*)

(*-----------------------------------------------------------------------------
 * 枚举: E_DL_SurgeState（归属本功能块，同文件发布，全库唯一定义）
 * 含义: 防喘振的工作相位。0 起步长 10。
 *-----------------------------------------------------------------------------*)
TYPE E_DL_SurgeState :
(
    eIdle        := 0,   // 待机：未使能 / Idle, disabled
    eNormal      := 10,  // 正常：流量高于危险线，阀关闭 / Normal, flow above the danger line, valve closed
    eRiskBlowoff := 20,  // 风险放空：流量低于危险线，阀快开 / Risk blowoff, valve fast open
    eRecovering  := 30,  // 恢复中：流量已越回差带，阀慢关 / Recovering, valve closing slowly
    eFault       := 99   // 故障：参数非法或输入非有限 / Fault, illegal parameter or non-finite input
);
END_TYPE

FUNCTION_BLOCK FB_DL_CompressorSurgeGuard
VAR_INPUT
    fSuctionPress   : REAL;                    // 吸入压力 [kPa abs]，须 > 0 / suction pressure [kPa abs], must be > 0
    fDischargePress : REAL;                    // 排出压力 [kPa abs] / discharge pressure [kPa abs]
    fFlow           : REAL;                    // 实测流量 [Nm3/h] / measured flow [Nm3/h]
    fFlowMinLine    : REAL := 500.0;           // 最小流量线 [Nm3/h]，须 > 0 / minimum flow line [Nm3/h], must be > 0
    fSurgeMargin    : REAL := 0.10;            // 危险线裕度 [倍]，须 > 0 / danger line margin [ratio], must be > 0
    fOpenRamp       : REAL := 20.0;            // 放空阀快开斜率 [%/s]，须 > 0 / blowoff fast-open ramp [%/s], must be > 0
    fCloseRamp      : REAL := 1.0;             // 放空阀慢关斜率 [%/s]，须 > 0 / blowoff slow-close ramp [%/s], must be > 0
    tConfirm        : TIME := T#200MS;         // 危险线确认时间 [ms] / danger line confirm time [ms]
    tSample         : TIME := T#100MS;         // 任务采样周期 [ms]，斜率换算用 / task sample period [ms], used by the ramps
    bEnable         : BOOL;                    // 使能 / enable
END_VAR
VAR_OUTPUT
    fBlowoffValve   : REAL;                    // 放空阀开度给定 [%]，范围 0~100 / blowoff valve opening setpoint [%], range 0~100
    bSurgeRisk      : BOOL;                    // 喘振风险（流量低于危险线，裸判据） / surge risk, the raw criterion
    bBlowoffActive  : BOOL;                    // 正在放空标志 / blowoff in progress flag
    fPressureRatio  : REAL;                    // 压比 = 排出/吸入 [倍] / pressure ratio, discharge over suction
    eErr            : UDINT;                   // 错误码，0 表示无错 / error code, 0 means no error
    bError          : BOOL;                    // 故障级标志，仅故障级错误置位 / fault-class flag, set only on fault-level codes
    bValid          : BOOL;                    // 输出可用标志 / outputs usable flag
END_VAR
VAR
    fbConfirm       : TON;                     // 危险线确认计时，段 6 无条件刷新 [ms] / danger line confirm timer
    fbRamp          : FB_DL_RateLimiter;       // 放空阀斜率限制子件（组合调用） / blowoff ramp subcomponent
    _eState         : E_DL_SurgeState := E_DL_SurgeState.eIdle; // 当前相位 / current phase
    _bInit          : BOOL := FALSE;           // 首扫标志，初值 FALSE 取非判定 / first-scan flag, tested negated
    _bFirstRamp     : BOOL := TRUE;            // 斜坡首次扫描跟踪标志（R36） / first-scan ramp tracking flag
    _bTrack         : BOOL := FALSE;           // 斜坡跟踪请求 / ramp tracking request
    _fTrackVal      : REAL;                    // 斜坡跟踪值 [%] / ramp tracking value [%]
    _bParamBad      : BOOL;                    // 参数非法标志 / illegal parameter flag
    _bFiniteBad     : BOOL;                    // 输入非有限标志 / non-finite input flag
    _bIllegal       : BOOL;                    // 非法状态标志 / illegal state flag
    _bRiskRaw       : BOOL;                    // 流量低于危险线（裸判据） / flow below the danger line, raw criterion
    _bRiskCfm       : BOOL;                    // 危险线确认条件（供定时器） / confirm condition for the timer
    _bRecovered     : BOOL;                    // 流量越出回差带 / flow recovered above the hysteresis band
    _bConfirmBreak  : BOOL;                    // 确认定时器断输入一拍标志 / confirm timer one-scan break
    _tConfirmUse    : TIME := T#200MS;         // 生效确认时间 [ms]，已钳位 / effective confirm time, clamped
    _fRatio         : REAL;                    // 压比 [倍] / pressure ratio
    _fRatioUse      : REAL := 1.0;             // 生效压比，夹到 ≥ 1 [倍] / effective ratio clamped to at least one
    _fDanger        : REAL;                    // 危险流量线 [Nm3/h] / danger flow line [Nm3/h]
    _fRecoverLine   : REAL;                    // 回差恢复线 [Nm3/h] / hysteresis recovery line [Nm3/h]
    _fTarget        : REAL;                    // 本拍目标阀位 [%] / target valve opening of this scan
    _fValveHeld     : REAL;                    // 末次阀位保持量 [%] / held valve opening [%]
    _fValvePrev     : REAL;                    // 上拍阀位（保持用，读子件前一拍输出） [%] / previous valve opening
    _fRampOut       : REAL;                    // 子件本拍输出 [%] / subcomponent output of this scan
END_VAR
VAR CONSTANT
    DL_PCT_MIN      : REAL := 0.0;             // 阀位下限 [%] / valve floor [%]
    DL_PCT_MAX      : REAL := 100.0;           // 阀位上限 [%] / valve ceiling [%]
    DL_VAL_LIM      : REAL := 1.0E30;          // 有限性判定的绝对值上限 [无量纲] / finiteness ceiling
    DL_RATIO_MIN    : REAL := 1.0;             // 压比可信下限 [倍]，低于 1 按 1 处理 / credible ratio floor, values below are clamped
    DL_SURGE_HYST   : REAL := 0.15;            // 恢复回差带 [倍]，禁裸数 / recovery hysteresis band [ratio], never a bare number
    DL_EPS          : REAL := 1.0E-6;          // 浮点比较容差 [%] / float comparison tolerance [%]
    DL_PARAM_MN     : REAL := 0.0;             // 参数下限，须严格大于 [无量纲] / parameter floor, must be strictly greater
    DL_CONF_MAX_MS  : DINT := 10000;           // 确认时间上限 [ms] / confirm time ceiling [ms]
    DL_TIME_ZERO    : TIME := T#0MS;           // 时间零值基准 [ms] / time zero reference
END_VAR

(*------------------------------------------------------------------------------
 * 段 1｜每拍预置（阀位与压比为保持量，在段 10 单点写入）
 *      Per-scan presets, the valve opening and the ratio are held and written once
 *-----------------------------------------------------------------------------*)
eErr           := 16#0000_0000;                // 错误码每拍重算 / error code recomputed every scan
bError         := FALSE;                       // 故障标志每拍重算 / fault flag recomputed every scan
bValid         := FALSE;                       // 可用标志每拍重算 / usable flag recomputed every scan
bSurgeRisk     := FALSE;                       // 风险位每拍重算 / risk flag recomputed every scan
bBlowoffActive := FALSE;                       // 放空动作位每拍重算 / blowoff active recomputed every scan
_bParamBad     := FALSE;                       // 参数非法标志预清零 / parameter flag pre-cleared
_bFiniteBad    := FALSE;                       // 非有限标志预清零 / non-finite flag pre-cleared
_bIllegal      := FALSE;                       // 非法状态标志预清零 / illegal state flag pre-cleared
_bRiskRaw      := FALSE;                       // 裸风险判据预置 FALSE / raw risk preset FALSE
_bRiskCfm      := FALSE;                       // 确认条件预置 FALSE / confirm condition preset FALSE
_bRecovered    := FALSE;                       // 恢复判据预置 FALSE / recovery preset FALSE
_bTrack        := FALSE;                       // 跟踪请求预置 FALSE / tracking request preset FALSE
_fTrackVal     := 0.0;                         // 跟踪值预置 0 [%] / tracking value preset to zero
_fRampOut      := 0.0;                         // 子件输出预置 0 [%] / subcomponent output preset to zero

(*------------------------------------------------------------------------------
 * 段 2｜首扫初始化（阀位从 0 起：放空阀失电关闭位）
 *      First-scan initialisation, the blowoff valve starts closed
 *-----------------------------------------------------------------------------*)
IF NOT _bInit THEN
    _eState     := E_DL_SurgeState.eIdle;      // 相位待机 / phase idle
    _fValveHeld := 0.0;                        // 阀位保持量 0 [%] / held valve opening zero
    _fRatio     := 0.0;                        // 压比保持量 0 [倍] / held ratio zero
    _bConfirmBreak := TRUE;                    // 确认计时从零开始 / confirm timer starts from zero
    _bFirstRamp := TRUE;                       // 斜坡首拍跟踪（R36） / ramp tracked on the first scan
    _bInit      := TRUE;                       // 首扫只做一次 / the first scan runs once
END_IF

(*------------------------------------------------------------------------------
 * 段 3｜参数闸门（含吸入压力 ≤ 0：压比无意义，按参数类处理）
 *      Parameter gate including a non-positive suction pressure, the ratio is meaningless then
 *-----------------------------------------------------------------------------*)
IF (fFlowMinLine <> fFlowMinLine) OR (ABS(fFlowMinLine) > DL_VAL_LIM) OR (fFlowMinLine <= DL_PARAM_MN) THEN
    _bParamBad := TRUE;                        // 最小流量线非法 / minimum flow line illegal
END_IF
IF (fSurgeMargin <> fSurgeMargin) OR (ABS(fSurgeMargin) > DL_VAL_LIM) OR (fSurgeMargin <= DL_PARAM_MN) THEN
    _bParamBad := TRUE;                        // 危险线裕度非法 / margin illegal
END_IF
IF (fOpenRamp <> fOpenRamp) OR (ABS(fOpenRamp) > DL_VAL_LIM) OR (fOpenRamp <= DL_PARAM_MN) THEN
    _bParamBad := TRUE;                        // 快开斜率非法 / fast-open ramp illegal
END_IF
IF (fCloseRamp <> fCloseRamp) OR (ABS(fCloseRamp) > DL_VAL_LIM) OR (fCloseRamp <= DL_PARAM_MN) THEN
    _bParamBad := TRUE;                        // 慢关斜率非法 / slow-close ramp illegal
END_IF
IF (fSuctionPress < -DL_VAL_LIM) OR (fSuctionPress > DL_VAL_LIM) THEN
    _bFiniteBad := TRUE;                       // 吸入压力非有限 / suction pressure non-finite
ELSIF fSuctionPress <= DL_PARAM_MN THEN
    _bParamBad := TRUE;                        // 吸入压力 ≤ 0：压比无意义 / non-positive suction, the ratio is meaningless
END_IF

(*------------------------------------------------------------------------------
 * 段 4｜其余输入的有限性闸门（区间判据同时拦 NaN 与 ±Inf）
 *      Finiteness gate for the remaining inputs
 *-----------------------------------------------------------------------------*)
IF (fDischargePress < -DL_VAL_LIM) OR (fDischargePress > DL_VAL_LIM) THEN
    _bFiniteBad := TRUE;                       // 排出压力非有限 / discharge pressure non-finite
END_IF
IF (fFlow < -DL_VAL_LIM) OR (fFlow > DL_VAL_LIM) THEN
    _bFiniteBad := TRUE;                       // 流量非有限 / flow non-finite
END_IF

(*------------------------------------------------------------------------------
 * 段 5｜压比与危险线（除零前置闸：吸入压力已确认 > 0，商前另设显式判据）
 *      Pressure ratio and danger line, the division is guarded twice
 *-----------------------------------------------------------------------------*)
IF (NOT _bFiniteBad) AND (NOT _bParamBad) THEN
    IF fSuctionPress > DL_PARAM_MN THEN
        _fRatio := fDischargePress / fSuctionPress; // 压比 [倍] / pressure ratio
    ELSE
        _fRatio := DL_RATIO_MIN;               // 结构性不可达（段 3 已拦），兜底为 1 / structurally unreachable fallback
    END_IF
    _fRatioUse := MAX(_fRatio, DL_RATIO_MIN);  // 夹到 ≥ 1：压比小于 1 的测量不可信 / clamp to at least one
    _fDanger   := fFlowMinLine * (1.0 + fSurgeMargin * (_fRatioUse - DL_RATIO_MIN)); // 危险流量线 [Nm3/h] / danger flow line
    _fRecoverLine := _fDanger * (1.0 + DL_SURGE_HYST); // 回差恢复线 [Nm3/h] / hysteresis recovery line
    _bRiskRaw  := (fFlow < _fDanger);          // 裸风险判据 [布尔] / raw risk criterion
    _bRecovered := (fFlow > _fRecoverLine);    // 越出回差带 [布尔] / recovered above the band
    _fRatio    := _fRatioUse;                  // 保持量取生效压比 / the held ratio is the effective one
END_IF

(*------------------------------------------------------------------------------
 * 段 6｜确认定时器无条件刷新（R40：CASE 之外每拍必调，转出相时断输入一拍）
 *      Confirm timer refreshed unconditionally outside the CASE
 *-----------------------------------------------------------------------------*)
_tConfirmUse := tConfirm;                      // 确认时间直取引脚 [ms] / confirm time taken from the pin
IF TIME_TO_DINT(_tConfirmUse) > DL_CONF_MAX_MS THEN
    _tConfirmUse := DINT_TO_TIME(DL_CONF_MAX_MS); // 超上限钳位（无专用码位，R90 不新开码） / clamped, no dedicated code
END_IF
IF TIME_TO_DINT(_tConfirmUse) < 0 THEN
    _tConfirmUse := DL_TIME_ZERO;              // 负时间结构性不可达，兜底为 0 / structurally unreachable fallback
END_IF

_bRiskCfm := bEnable AND (NOT _bParamBad) AND (NOT _bFiniteBad) AND _bRiskRaw; // 确认条件

fbConfirm(IN := _bRiskCfm AND (NOT _bConfirmBreak), PT := _tConfirmUse); // 危险线确认计时无条件刷新
_bConfirmBreak := FALSE;                       // 断输入拍在调用后自清（R40 自清位置） / break self-cleared after the call

(*------------------------------------------------------------------------------
 * 段 7｜相位机（只做迁移；阀位与码位在段 9/10 处理）
 *      Phase machine, transitions only
 *-----------------------------------------------------------------------------*)
CASE _eState OF

    E_DL_SurgeState.eIdle:                     // 待机：参数合法、输入有限且使能即进入
        IF _bParamBad OR _bFiniteBad THEN
            _eState := E_DL_SurgeState.eFault; // 原因未消失，转故障 / the cause persists
        ELSIF bEnable THEN
            IF _bRiskRaw AND fbConfirm.Q THEN
                _eState := E_DL_SurgeState.eRiskBlowoff; // 已确认风险，直接进放空 / confirmed risk
            ELSE
                _eState := E_DL_SurgeState.eNormal; // 进正常相 / enter the normal phase
            END_IF
        END_IF

    E_DL_SurgeState.eNormal:                   // 正常：流量低于危险线并确认即放空
        IF _bParamBad OR _bFiniteBad THEN
            _eState := E_DL_SurgeState.eFault; // 转故障 / go to fault
        ELSIF NOT bEnable THEN
            _eState := E_DL_SurgeState.eIdle;  // 失能回待机 / disabled, back to idle
        ELSIF _bRiskRaw AND fbConfirm.Q THEN
            _eState := E_DL_SurgeState.eRiskBlowoff; // 风险确认，进放空 / risk confirmed, blow off
            _bConfirmBreak := TRUE;            // 换相后确认计时重启 / restart the confirm timer across the phase change
        END_IF

    E_DL_SurgeState.eRiskBlowoff:              // 风险放空：必须经恢复相，不得被 eNormal 直接抢占
        IF _bParamBad OR _bFiniteBad THEN
            _eState := E_DL_SurgeState.eFault; // 转故障 / go to fault
        ELSIF NOT bEnable THEN
            _eState := E_DL_SurgeState.eIdle;  // 失能回待机 / disabled, back to idle
        ELSIF _bRecovered THEN
            _eState := E_DL_SurgeState.eRecovering; // 越出回差带，进慢关相 / recovered, start closing slowly
        END_IF

    E_DL_SurgeState.eRecovering:               // 恢复中：再次跌破危险线则回放空，阀关到 0 才回正常
        IF _bParamBad OR _bFiniteBad THEN
            _eState := E_DL_SurgeState.eFault; // 转故障 / go to fault
        ELSIF NOT bEnable THEN
            _eState := E_DL_SurgeState.eIdle;  // 失能回待机 / disabled, back to idle
        ELSIF _bRiskRaw THEN
            _eState := E_DL_SurgeState.eRiskBlowoff; // 再次跌破危险线，回放空 / below the danger line again
        ELSIF _fValvePrev <= DL_PCT_MIN + DL_EPS THEN
            _eState := E_DL_SurgeState.eNormal; // 阀已关到 0，回正常 / the valve is closed, back to normal
        END_IF

    E_DL_SurgeState.eFault:                    // 故障：原因消失即自动恢复（本件无复位引脚）
        IF NOT bEnable THEN
            _eState := E_DL_SurgeState.eIdle;  // 失能回待机 / disabled, back to idle
        ELSIF (NOT _bParamBad) AND (NOT _bFiniteBad) THEN
            _eState := E_DL_SurgeState.eNormal; // 原因消失自动回正常 / cause cleared, resume
        END_IF

    ELSE
        _bIllegal := TRUE;                     // 标记非法状态 / flag the illegal state
        _eState   := E_DL_SurgeState.eFault;   // 回故障态 / back to the fault state
END_CASE

(*------------------------------------------------------------------------------
 * 段 8｜目标阀位（两条安全方向相反的规则在此并列，不得只做其一）
 *      Target valve opening, the two opposite safety rules live side by side here
 *-----------------------------------------------------------------------------*)
_fValvePrev := fbRamp.fOut;                    // 先读子件上一拍输出 [%] / read the subcomponent output first

IF _bIllegal OR _bParamBad THEN
    _fTarget := DL_PCT_MAX;                    // 参数/状态非法：阀全开（宁可放空不可喘振） [%] / illegal, full open
    eErr     := 16#0005_030B;                  // 故障级：参数非法，阀全开 / fault: illegal parameter, valve fully open
    bError   := TRUE;                          // 置故障标志 / raise the fault flag
ELSIF _bFiniteBad THEN
    _fTarget := _fValvePrev;                   // 非有限：目标 = 当前阀位，即保持（坏值不得关阀） [%] / hold the valve
    eErr     := 16#0005_030C;                  // 故障级：输入非有限，保持末次阀位 / fault: non-finite input, valve held
    bError   := TRUE;                          // 置故障标志 / raise the fault flag
ELSIF NOT bEnable THEN
    _fTarget := DL_PCT_MIN;                    // 失能：慢关到 0（走慢关斜率，不阶跃） [%] / disabled, close slowly
    _bConfirmBreak := TRUE;                    // 失能时确认计时重启 / restart the confirm timer
ELSIF _eState = E_DL_SurgeState.eRiskBlowoff THEN
    _fTarget := DL_PCT_MAX;                    // 风险放空：阀全开（由快开斜率跟随） [%] / risk blowoff, full open
    eErr     := 16#0005_01DA;                  // 信息级：流量低于危险线已开放空阀 / informational: blowoff opened
ELSIF _eState = E_DL_SurgeState.eRecovering THEN
    _fTarget := DL_PCT_MIN;                    // 恢复中：慢关（由慢关斜率跟随） [%] / recovering, close slowly
    eErr     := 16#0005_01DB;                  // 信息级：已退出放空 / informational: leaving blowoff
ELSE
    _fTarget := DL_PCT_MIN;                    // 正常：阀关闭 [%] / normal, valve closed
END_IF

(*------------------------------------------------------------------------------
 * 段 9｜斜坡组合调用（快开慢关各用一支斜率，跟踪注入按 R36 手算首拍）
 *      Ramp composition, fast open and slow close, tracking injected per R36
 *-----------------------------------------------------------------------------*)
_bTrack   := _bFiniteBad OR _bFirstRamp;       // 非有限保持与首次扫描都走跟踪，避免阶跃 / hold and first scan are tracked
_fTrackVal := _fValvePrev;                     // 跟踪值 = 当前阀位 [%] / tracking value is the current opening
IF _bFirstRamp THEN
    _fTrackVal := _fValveHeld;                 // 首拍跟踪到保持量（初始为 0） [%] / first scan tracks the held value
END_IF

fbRamp(bEnable     := TRUE,                    // 子件恒使能：斜率限制始终生效 / always enabled, the ramp always applies
       fIn         := _fTarget,                // 目标阀位 [%] / target opening
       fRateUp      := fOpenRamp,              // 快开斜率 [%/s] / fast-open ramp
       fRateDown    := fCloseRamp,             // 慢关斜率 [%/s] / slow-close ramp
       bTrack       := _bTrack,                // 跟踪请求 / tracking request
       fTrackValue  := _fTrackVal,             // 跟踪值 [%] / tracking value
       tSampleTime  := tSample);               // 采样周期 [ms] / sample period
_fRampOut   := fbRamp.fOut;                    // 取子件输出 [%] / take the subcomponent output
_bFirstRamp := FALSE;                          // 首拍跟踪只做一次 / first-scan tracking runs once

(*------------------------------------------------------------------------------
 * 段 10｜输出单点写入与可用性仲裁
 *      Single write point of the outputs and the usability arbitration
 *-----------------------------------------------------------------------------*)
_fRampOut   := LIMIT(DL_PCT_MIN, _fRampOut, DL_PCT_MAX); // 子件输出再钳一次（防御纵深） [%] / clamped again, defense in depth
_fValveHeld := _fRampOut;                      // 阀位保持量跟进 [%] / the held opening follows
fBlowoffValve := _fRampOut;                    // 阀位出口 [%] / valve opening outlet
fPressureRatio := _fRatio;                     // 压比出口 [倍] / pressure ratio outlet
bSurgeRisk    := _bRiskRaw;                    // 风险位保持可观测（失能亦然） / the risk stays observable even when disabled
bBlowoffActive := (_eState = E_DL_SurgeState.eRiskBlowoff); // 正在放空：仅风险相为真 / blowoff active in the risk phase only

IF bError THEN
    bValid := FALSE;                           // 故障级：输出不可用 / fault: outputs unusable
ELSIF NOT bEnable THEN
    bValid := FALSE;                           // 失能：输出不可用（阀位仍按慢关下落） / disabled: unusable, the valve still closes
ELSIF _bIllegal THEN
    bValid := FALSE;                           // 非法状态：输出不可用 / illegal state: unusable
ELSE
    bValid := TRUE;                            // 输出可用 / outputs usable
END_IF

END_FUNCTION_BLOCK
